(* IEC 61131-3 sources: JingjiangArm/moonboxpro_arm_8.4/Application/Application/任务列表/CommTask/COMM_DIAMONDS/Input_Output, 7 files *)

(* ---- KS_CheckStationOnLine_.st ---- *)
(*@CES
Name=KS_CheckStationOnLine_
Type=FunctionBlock
TypeGuid=6f9dac99-8de1-4efc-8465-68ac443b7d08
Guid=c5e0cdd1-19ab-4cb0-a985-998ee908852c
HasDeclaration=True
HasImplementation=True
*)
{DECLARATION}
FUNCTION KS_CheckStationOnLine_ : BOOL
VAR_INPUT
	i_iSid : INT;
	i_iStationNum : INT;
	i_paiStationId_List : POINTER TO ARRAY [1..128] OF INT;
END_VAR
VAR
	iN : INT;
	xResult : BOOL;
END_VAR

{IMPLEMENTATION}
xResult := FALSE;

FOR iN := 1 TO i_iStationNum BY 1 DO
	IF i_iSid = i_paiStationId_List^[iN] THEN
		xResult := TRUE;
		EXIT;
	END_IF
END_FOR

KS_CheckStationOnLine_ := xResult;

(* ---- KS_Solve_Ver.st ---- *)
(*@CES
Name=KS_Solve_Ver
Type=FunctionBlock
TypeGuid=6f9dac99-8de1-4efc-8465-68ac443b7d08
Guid=eb7c1164-08c4-4977-9280-cbaed44442c1
HasDeclaration=True
HasImplementation=True
*)
{DECLARATION}
FUNCTION KS_Solve_Ver : BOOL(*版本号解析*)
VAR_INPUT
	i_sVersion: STRING;(*版本号*)
	i_pdwYMD: POINTER TO DWORD;
	i_pdwHMS: POINTER TO DWORD;
	i_pdwVer: POINTER TO DWORD;
END_VAR
VAR
END_VAR

{IMPLEMENTATION}
IF i_pdwYMD<>0 AND i_pdwHMS<>0 AND i_pdwVer<>0 THEN

END_IF

(* ---- KS_FB_DIAMONDS_Input.st ---- *)
(*@CES
Name=KS_FB_DIAMONDS_Input
Type=FunctionBlock
TypeGuid=6f9dac99-8de1-4efc-8465-68ac443b7d08
Guid=1e0a50ec-9206-4692-bb5f-e2a5b8087577
HasDeclaration=True
HasImplementation=True
*)
{DECLARATION}
FUNCTION_BLOCK KS_FB_DIAMONDS_Input
VAR_INPUT
	i_xEn: BOOL;
	i_pstStSysParam: POINTER TO StSysParam;
	i_pstStParam_Diamonds_Wr: POINTER TO StParam_Diamonds_Wr;
	i_pstStParam_Diamonds_WrRd: POINTER TO StParam_Diamonds_WrRd;
	i_pstStWrRd_SysCfg: POINTER TO StWrRd_SysCfg;
	i_pstStSysCfgStruct: POINTER TO StSysCfgStruct;
	i_pastStGetMotionSts: POINTER TO ARRAY [1..MAX_STATION_NUM] OF StGetMotionSts;

END_VAR
VAR_OUTPUT
	o_xEn: BOOL;
	o_iErNo: INT;
END_VAR
VAR
	pstStParam_Diamonds_Wr_SysSts : POINTER TO StParam_Diamonds_Wr_SysSts;
	pstStParam_Diamonds_Wr_RdSam : POINTER TO StParam_Diamonds_Wr_RdSam;
	pastStParam_Diamonds_Wr_Err : POINTER TO ARRAY [1..MAX_UNIT_NUM] OF StParam_Diamonds_Wr_Err;
	pastStParam_Diamonds_Wr_RunSts : POINTER TO ARRAY [1..MAX_STATION_NUM] OF StParam_Diamonds_Wr_RunSts;
	iGrp: INT;
	iUnitId: INT;
	byCurSignal_RGB: BYTE;
	abySignalFlag: ARRAY [1..4] OF BYTE;
	iIndex:INT:= 1;
	iN: INT;
	iJ: INT;
	iK: INT;

	abyLastIndex: ARRAY [1..MAX_UNIT_NUM] OF BYTE;
	iAxisId_If: INT;
	iAxisId_Of: INT;
	iGrpId_Uw: INT;
	iGrpId_Rw: INT;
	fbKS_FB_DIAMONDS_SysCfg_WrRd: KS_FB_DIAMONDS_SysCfg_WrRd;
	iMachanicalTypeId: INT;

	astStParam_Diamonds_Wr_RunSts : ARRAY [1..MAX_STATION_NUM] OF StParam_Diamonds_Wr_RunSts;
	iNumIndex: INT:=0;
	iAxisId_T: INT;
	iTypeId_T: INT;
	iUnitId_T: INT;
	iCoreId_T: INT;
	iGroupId_T: INT;
	iAdjAxisId_T: INT;

END_VAR

{IMPLEMENTATION}
o_xEn:= i_xEn;
o_iErNo:= 0;
IF i_xEn THEN
	IF i_pstStSysParam<>0 AND
		i_pstStParam_Diamonds_Wr<>0 AND
		i_pstStParam_Diamonds_WrRd<>0 THEN
		pstStParam_Diamonds_Wr_SysSts:= ADR(i_pstStParam_Diamonds_Wr^.stStParam_Diamonds_Wr_SysSts);
		pstStParam_Diamonds_Wr_RdSam:= ADR(i_pstStParam_Diamonds_Wr^.stStParam_Diamonds_Wr_RdSam);
		pastStParam_Diamonds_Wr_Err:= ADR(i_pstStParam_Diamonds_Wr^.astStParam_Diamonds_Wr_Err);
		pastStParam_Diamonds_Wr_RunSts:= ADR(i_pstStParam_Diamonds_Wr^.astStParam_Diamonds_Wr_RunSts);

		Action_Input_Wr();
(*2025.8.6.195943*)
//2026.5.29.145241		Action_Input_WrRd();

		o_iErNo:= 1;
	ELSE
		o_iErNo:= -2;
	END_IF
ELSE
	o_iErNo:= -1;
END_IF

(* ---- KS_FB_DIAMONDS_Input_WRRD.st ---- *)
(*@CES
Name=KS_FB_DIAMONDS_Input_WRRD
Type=FunctionBlock
TypeGuid=6f9dac99-8de1-4efc-8465-68ac443b7d08
Guid=edee9bc0-245c-42df-bd06-57a10449e106
HasDeclaration=True
HasImplementation=True
*)
{DECLARATION}
FUNCTION_BLOCK KS_FB_DIAMONDS_Input_WRRD
VAR_INPUT
	i_xEn: BOOL;
	i_pstStSysParam: POINTER TO StSysParam;
	i_pstStParam_Diamonds_WrRd: POINTER TO StParam_Diamonds_WrRd;
	i_pstStWrRd_SysCfg: POINTER TO StWrRd_SysCfg;
	i_pstStSysCfgStruct: POINTER TO StSysCfgStruct;

END_VAR
VAR_OUTPUT
	o_xEn: BOOL;
	o_iErNo: INT;
END_VAR
VAR
	iGrp: INT;
	iUnitId: INT;
	byCurSignal_RGB: BYTE;
	abySignalFlag: ARRAY [1..4] OF BYTE;
	iIndex:INT:= 1;
	iN: INT;
	iJ: INT;
	iK: INT;

	abyLastIndex: ARRAY [1..MAX_UNIT_NUM] OF BYTE;
	iAxisId_If: INT;
	iAxisId_Of: INT;
	iGrpId_Uw: INT;
	iGrpId_Rw: INT;
	fbKS_FB_DIAMONDS_SysCfg_WrRd: KS_FB_DIAMONDS_SysCfg_WrRd;
	iMachanicalTypeId: INT;
	iMachanicalTypeId_Tmp: INT;

END_VAR

{IMPLEMENTATION}
(*整机参数|2025.08.06.203301*)
	i_pstStParam_Diamonds_WrRd^.iCustomerId 													:= i_pstStSysParam^.stStSysParam_Save.iCustomerId;									(*客户ID*)
	i_pstStParam_Diamonds_WrRd^.dwEquipmentProf 												:= i_pstStSysParam^.stStSysParam_Save.dwEquipmentProf;								(*设备描述*)
	i_pstStParam_Diamonds_WrRd^.iUnitMaxNum 													:= i_pstStSysParam^.stStSysParam_Save.iUnitMaxNum;												(*最大色组数*)
	i_pstStParam_Diamonds_WrRd^.iCurveViewMaxRange 												:= i_pstStSysParam^.stStSysParam_Save.iCurveViewMaxRange;							(*误差曲线量程上限*)
	i_pstStParam_Diamonds_WrRd^.iTitleTextHeight 												:= i_pstStSysParam^.stStSysParam_Save.iTitleTextHeight;								(*标题字体高度*)
	i_pstStParam_Diamonds_WrRd^.iEntryTextHeight 												:= i_pstStSysParam^.stStSysParam_Save.iEntryTextHeight;								(*输入框字体高度*)
	i_pstStParam_Diamonds_WrRd^.iLabelTextHeight 												:= i_pstStSysParam^.stStSysParam_Save.iLabelTextHeight;								(*标签字体高度*)
	i_pstStParam_Diamonds_WrRd^.iButtonTextHeight 												:= i_pstStSysParam^.stStSysParam_Save.iButtonTextHeight ;							(*按钮字体高度*)
	i_pstStParam_Diamonds_WrRd^.iMessageTextHeight 												:= i_pstStSysParam^.stStSysParam_Save.iMessageTextHeight;							(*消息字体高度*)
	i_pstStParam_Diamonds_WrRd^.byLanguageId 													:= i_pstStSysParam^.stStSysParam_Save.byLanguageId;									(*语言设置*)
	i_pstStParam_Diamonds_WrRd^.byMinutes_ScrSaver 												:= i_pstStSysParam^.stStSysParam_Save.byMinutes_ScrSaver;							(*屏保延时*)
	i_pstStParam_Diamonds_WrRd^.wMachineArchitectureRef 										:= i_pstStSysParam^.stStSysParam_Save.wMachineArchitectureRef;						(*机器架构描述*)
	i_pstStParam_Diamonds_WrRd^.iPromptMsgId 													:= i_pstStSysParam^.stStSysParam_Save.iPromptMsgId;									(*提示信息ID（报警代码）*)
	i_pstStParam_Diamonds_WrRd^.byHorzCtlMode 													:= i_pstStSysParam^.stStSysParam_Save.byHorzCtlMode;								(*横向控制方式-同步-步进-伺服*)
	i_pstStParam_Diamonds_WrRd^.byCheckTimeToTips_BrakeResistance 								:= i_pstStSysParam^.stStSysParam_Save.byCheckTimeToTips_BrakeResistance;			(*制动电阻访问超限提示时间*)
	i_pstStParam_Diamonds_WrRd^.byCheckTimeToEStop_BrakeResistance 								:= i_pstStSysParam^.stStSysParam_Save.byCheckTimeToEStop_BrakeResistance;			(*制动电阻访问超限急停时间*)
	i_pstStParam_Diamonds_WrRd^.byAccessTimes_BrakeResistance 									:= i_pstStSysParam^.stStSysParam_Save.byAccessTimes_BrakeResistance;				(*制动电阻报警限制*)
	i_pstStParam_Diamonds_WrRd^.byAlarmHold_VOL_Uw 												:= i_pstStSysParam^.stStSysParam_Save.byAlarmHold_VOL_Uw;							(*放料没料响应时间*)
	i_pstStParam_Diamonds_WrRd^.byAlarmHold_PrnLength 											:= i_pstStSysParam^.stStSysParam_Save.byAlarmHold_PrnLength;						(*收料印长报警响应时间*)
	i_pstStParam_Diamonds_WrRd^.byHeatingOutWay_III 											:= i_pstStSysParam^.stStSysParam_Save.byHeatingOutWay_III;							(*三档调整方式-只调最低档、只调最高档、三档同时调*)
	i_pstStParam_Diamonds_WrRd^.byHeatingMode 													:= i_pstStSysParam^.stStSysParam_Save.byHeatingMode;								(*温控设置方式切换*)
	i_pstStParam_Diamonds_WrRd^.rOpenThr_Ele 													:= i_pstStSysParam^.stStSysParam_Save.rOpenThr_Ele;									(*电加热开启*)
	i_pstStParam_Diamonds_WrRd^.rCloseThr_Ele 													:= i_pstStSysParam^.stStSysParam_Save.rCloseThr_Ele;								(*电加热关闭*)
	i_pstStParam_Diamonds_WrRd^.rDealValue_Water 												:= i_pstStSysParam^.stStSysParam_Save.rDealValue_Water;								(*水加热死区*)
	i_pstStParam_Diamonds_WrRd^.iMaxOutValue 													:= i_pstStSysParam^.stStSysParam_Save.iMaxOutValue;									(*最大输出*)
	i_pstStParam_Diamonds_WrRd^.iHeatingDebugValue_Water 										:= i_pstStSysParam^.stStSysParam_Save.iHeatingDebugValue_Water;						(*测试开度*)
	i_pstStParam_Diamonds_WrRd^.rKp 															:= i_pstStSysParam^.stStSysParam_Save.rKp;											(*KP*)
	i_pstStParam_Diamonds_WrRd^.rKi 															:= i_pstStSysParam^.stStSysParam_Save.rKi;											(*KI*)
	i_pstStParam_Diamonds_WrRd^.rKd 															:= i_pstStSysParam^.stStSysParam_Save.rKd;											(*Kd*)
	i_pstStParam_Diamonds_WrRd^.iTime_Thres_Water 												:= i_pstStSysParam^.stStSysParam_Save.iTime_Thres_Water;							(*阀门打开时间*)
	i_pstStParam_Diamonds_WrRd^.iCofe_TempCtl_30 												:= i_pstStSysParam^.stStSysParam_Save.iCofe_TempCtl_30;								(*控制阈值1*)
	i_pstStParam_Diamonds_WrRd^.iCofe_TempCtl_30_10 											:= i_pstStSysParam^.stStSysParam_Save.iCofe_TempCtl_30_10;							(*控制阈值2*)
	i_pstStParam_Diamonds_WrRd^.iCofe_TempCtl_10_5 												:= i_pstStSysParam^.stStSysParam_Save.iCofe_TempCtl_10_5;							(*控制阈值3*)
	i_pstStParam_Diamonds_WrRd^.iCofe_TempCtl_5 												:= i_pstStSysParam^.stStSysParam_Save.iCofe_TempCtl_5;								(*控制阈值4*)
	i_pstStParam_Diamonds_WrRd^.iWaterValue_Threshold 											:= i_pstStSysParam^.stStSysParam_Save.iWaterValue_Threshold;						(*水电阈值*)
	i_pstStParam_Diamonds_WrRd^.uiInitDiam_Uw 													:= i_pstStSysParam^.stStSysParam_Save.uiInitDiam_Uw;								(*放料初始卷径*)
	i_pstStParam_Diamonds_WrRd^.uiInitDiam_Rw 													:= i_pstStSysParam^.stStSysParam_Save.uiInitDiam_Rw;								(*收料初始卷径*)
	i_pstStParam_Diamonds_WrRd^.diStepDriveDebugPulse 											:= i_pstStSysParam^.stStSysParam_Save.diStepDriveDebugPulse;						(*测试脉冲数*)
	i_pstStParam_Diamonds_WrRd^.rStepDriveDebugPulse_PosAct 									:= i_pstStSysParam^.stStSysParam_Save.rStepDriveDebugPulse_PosAct;					(*测试距离*)
	i_pstStParam_Diamonds_WrRd^.iStepDriveDebugNum 												:= i_pstStSysParam^.stStSysParam_Save.iStepDriveDebugNum;							(*测试色组号*)
	i_pstStParam_Diamonds_WrRd^.rStepDrivePosPPulse 											:= i_pstStSysParam^.stStSysParam_Save.rStepDrivePosPPulse;							(*单位脉冲距离*)
	i_pstStParam_Diamonds_WrRd^.iStepDrivePulsePRev 											:= i_pstStSysParam^.stStSysParam_Save.iStepDrivePulsePRev;							(*每圈脉冲数*)
	i_pstStParam_Diamonds_WrRd^.iStepDriveSa_Vel 												:= i_pstStSysParam^.stStSysParam_Save.iStepDriveSa_Vel;								(*启动速度*)
	i_pstStParam_Diamonds_WrRd^.iStepDrivePreReg_Vel 											:= i_pstStSysParam^.stStSysParam_Save.iStepDrivePreReg_Vel;							(*预套准速度*)
	i_pstStParam_Diamonds_WrRd^.iStepDriveManu_Vel 												:= i_pstStSysParam^.stStSysParam_Save.iStepDriveManu_Vel;							(*手动低速*)
	i_pstStParam_Diamonds_WrRd^.iStepDriveManu_Vel_Fast 										:= i_pstStSysParam^.stStSysParam_Save.iStepDriveManu_Vel_Fast;						(*手动高速*)
	i_pstStParam_Diamonds_WrRd^.iStepDriveAuto_Vel 												:= i_pstStSysParam^.stStSysParam_Save.iStepDriveAuto_Vel;							(*自动速度*)
	i_pstStParam_Diamonds_WrRd^.iStepDriveAccTime 												:= i_pstStSysParam^.stStSysParam_Save.iStepDriveAccTime;							(*升速时间*)
	i_pstStParam_Diamonds_WrRd^.rHz_MainExhaust_ManuallySet 									:= i_pstStSysParam^.stStSysParam_Save.rHz_MainExhaust_ManuallySet;					(*主排风设定频率*)
	i_pstStParam_Diamonds_WrRd^.byFreq_I_ExhaustAir 											:= i_pstStSysParam^.stStSysParam_Save.byFreq_I_ExhaustAir;							(*排风一档频率*)
	i_pstStParam_Diamonds_WrRd^.byFreq_II_ExhaustAir 											:= i_pstStSysParam^.stStSysParam_Save.byFreq_II_ExhaustAir;							(*排风二档频率*)
	i_pstStParam_Diamonds_WrRd^.byFreq_III_ExhaustAir 											:= i_pstStSysParam^.stStSysParam_Save.byFreq_III_ExhaustAir;						(*排风三档频率*)
	(*待补充-开始|2025.08.06.210116*)
	i_pstStParam_Diamonds_WrRd^.stBitStWrRd_Switch_Machine.xSwitch_PreHotEn_Print				:= i_pstStSysParam^.stStSysParam_Save.xSwitch_PreHotEn_Print				;(*预热印刷激活开关*)
	i_pstStParam_Diamonds_WrRd^.stBitStWrRd_Switch_Machine.xSwitch_ExhAir_Limit_HotWind			:= i_pstStSysParam^.stStSysParam_Save.xSwitch_ExhAir_Limit_HotWind			;(*排风限制热风开关*)
	i_pstStParam_Diamonds_WrRd^.stBitStWrRd_Switch_Machine.xSwitch_ExhAir_Limit_Run				:= i_pstStSysParam^.stStSysParam_Save.xSwitch_ExhAir_Limit_Run				;(*排风限制开机开关*)
	i_pstStParam_Diamonds_WrRd^.stBitStWrRd_Switch_Machine.xSwitch_CommEn_WatchDevice_Tcp		:= i_pstStSysParam^.stStSysParam_Save.xSwitch_CommEn_WatchDevice_Tcp		;(*TCP-外部监控设备开关*)
	i_pstStParam_Diamonds_WrRd^.stBitStWrRd_Switch_Machine.xSwitch_CommEn_WatchDevice_485		:= i_pstStSysParam^.stStSysParam_Save.xSwitch_CommEn_WatchDevice_485		;(*485-外部监控设备开关*)
	i_pstStParam_Diamonds_WrRd^.stBitStWrRd_Switch_Machine.xSwitch_CommEn_1U_485				:= i_pstStSysParam^.stStSysParam_Save.xSwitch_CommEn_1U_485				    ;(*1色人机通讯开关*)
	i_pstStParam_Diamonds_WrRd^.stBitStWrRd_Switch_Machine.xSwitch_CommEn_485					:= i_pstStSysParam^.stStSysParam_Save.xSwitch_CommEn_485					;(*485通讯开关*)
	i_pstStParam_Diamonds_WrRd^.stBitStWrRd_Switch_Machine.xSwitch_CommEn_485_Exh				:= i_pstStSysParam^.stStSysParam_Save.xSwitch_CommEn_485_Exh				;(*排风485通讯开关*)
	i_pstStParam_Diamonds_WrRd^.stBitStWrRd_Switch_Machine.xSwitch_CommEn_485_Scraper			:= i_pstStSysParam^.stStSysParam_Save.xSwitch_CommEn_485_Scraper			;(*刮刀485通讯开关*)
	i_pstStParam_Diamonds_WrRd^.stBitStWrRd_Switch_Machine.xSwitch_CommEn_485_InkRoller			:= i_pstStSysParam^.stStSysParam_Save.xSwitch_CommEn_485_InkRoller			;(*递墨辊485通讯开关*)
	i_pstStParam_Diamonds_WrRd^.stBitStWrRd_Switch_Machine.xSwitch_CommEn_485_HotWind			:= i_pstStSysParam^.stStSysParam_Save.xSwitch_CommEn_485_HotWind			;(*热风485通讯开关*)
	i_pstStParam_Diamonds_WrRd^.stBitStWrRd_Switch_Machine.xSwitch_ArcIntensityBtn_Hmi			:= i_pstStSysParam^.stStSysParam_Save.xSwitch_ArcIntensityBtn_Hmi			;(*手动调节随速度走开关*)
	i_pstStParam_Diamonds_WrRd^.stBitStWrRd_Switch_Machine.xSwitch_PrnRatioIndividual_Setting	:= i_pstStSysParam^.stStSysParam_Save.xSwitch_PrnRatioIndividual_Setting	;(*色组版辊减速比单独设置开关*)
	i_pstStParam_Diamonds_WrRd^.stBitStWrRd_Switch_Machine.xSwitch_NetRatioIndividual_Setting	:= i_pstStSysParam^.stStSysParam_Save.xSwitch_NetRatioIndividual_Setting	;(*色组网辊减速比单独设置开关*)
	i_pstStParam_Diamonds_WrRd^.stBitStWrRd_Switch_Machine.xSwitch_BottomRatioIndividual_Setting:= i_pstStSysParam^.stStSysParam_Save.xSwitch_BottomRatioIndividual_Setting ;(*色组底辊减速比单独设置开关*)
	i_pstStParam_Diamonds_WrRd^.stBitStWrRd_Switch_Machine.xSwitch_StepDriveDebugRun			:= i_pstStSysParam^.stStSysParam_Save.xSwitch_StepDriveDebugRun			    ;(*横向步进电机测试执行开关*)

	i_pstStParam_Diamonds_WrRd^.stBitStWrRd_Switch_Machine.xSetProPointEn					 := i_pstStSysParam^.stStSysParam_Save.xSetProPointEn					;
	i_pstStParam_Diamonds_WrRd^.stBitStWrRd_Switch_Machine.xUseMaxTimeAsSBegin_InLowSpeed    := i_pstStSysParam^.stStSysParam_Save.xUseMaxTimeAsSBegin_InLowSpeed	;
	i_pstStParam_Diamonds_WrRd^.stBitStWrRd_Switch_Machine.xPseudoRandomEn                   := i_pstStSysParam^.stStSysParam_Save.xPseudoRandomEn               	;
	i_pstStParam_Diamonds_WrRd^.stBitStWrRd_Switch_Machine.xPseudoRandomStart                := i_pstStSysParam^.stStSysParam_Save.xPseudoRandomStart            	;
	i_pstStParam_Diamonds_WrRd^.stBitStWrRd_Switch_Machine.xEn_RevLimit                      := i_pstStSysParam^.stStSysParam_Save.xEn_RevLimit                  	;
	i_pstStParam_Diamonds_WrRd^.stBitStWrRd_Switch_Machine.xSaveFineSampleData_ToArc         := i_pstStSysParam^.stStSysParam_Save.xSaveFineSampleData_ToArc     	;
	i_pstStParam_Diamonds_WrRd^.stBitStWrRd_Switch_Machine.xReqSetLedFunc                    := i_pstStSysParam^.stStSysParam_Save.xReqSetLedFunc                	;
	i_pstStParam_Diamonds_WrRd^.stBitStWrRd_Switch_Machine.xSetHmiResolution                 := i_pstStSysParam^.stStSysParam_Save.xSetHmiResolution             	;
	i_pstStParam_Diamonds_WrRd^.stBitStWrRd_Switch_Machine.xPopupWindowVisible               := i_pstStSysParam^.stStSysParam_Save.xPopupWindowVisible           	;
	i_pstStParam_Diamonds_WrRd^.stBitStWrRd_Switch_Machine.xInitArcErr_AjdImmediately        := i_pstStSysParam^.stStSysParam_Save.xInitArcErr_AjdImmediately    	;
	i_pstStParam_Diamonds_WrRd^.stBitStWrRd_Switch_Machine.xPhaseAutoRecoveryEn              := i_pstStSysParam^.stStSysParam_Save.xPhaseAutoRecoveryEn          	;
	i_pstStParam_Diamonds_WrRd^.stBitStWrRd_Switch_Machine.xKeepServo_PreRegisterDne         := i_pstStSysParam^.stStSysParam_Save.xKeepServo_PreRegisterDne     	;
	i_pstStParam_Diamonds_WrRd^.stBitStWrRd_Switch_Machine.xUseIfVel_Uw                      := i_pstStSysParam^.stStSysParam_Save.xUseIfVel_Uw                  	;
	i_pstStParam_Diamonds_WrRd^.stBitStWrRd_Switch_Machine.xKeepServo_Stop                   := i_pstStSysParam^.stStSysParam_Save.xKeepServo_Stop               	;
	i_pstStParam_Diamonds_WrRd^.stBitStWrRd_Switch_Machine.xAxisPrfVelEn                     := i_pstStSysParam^.stStSysParam_Save.xAxisPrfVelEn                 	;
	i_pstStParam_Diamonds_WrRd^.stBitStWrRd_Switch_Machine.xUseGc_PID_2025                   := i_pstStSysParam^.stStSysParam_Save.xUseGc_PID_2025               	;
	i_pstStParam_Diamonds_WrRd^.stBitStWrRd_Switch_Machine.xFlag_Follow_1U_Double_V          := i_pstStSysParam^.stStSysParam_Save.xFlag_Follow_1U_Double_V      	;
	i_pstStParam_Diamonds_WrRd^.stBitStWrRd_Switch_Machine.xArcErrCorrectIsRev_V             := i_pstStSysParam^.stStSysParam_Save.xArcErrCorrectIsRev_V         	;
	i_pstStParam_Diamonds_WrRd^.stBitStWrRd_Switch_Machine.xAutoSetSampleType                := i_pstStSysParam^.stStSysParam_Save.xAutoSetSampleType            	;
	i_pstStParam_Diamonds_WrRd^.stBitStWrRd_Switch_Machine.xGetSampleTypeBtn                 := i_pstStSysParam^.stStSysParam_Save.xGetSampleTypeBtn             	;
	i_pstStParam_Diamonds_WrRd^.stBitStWrRd_Switch_Machine.xAutoSetArcCtlWay                 := i_pstStSysParam^.stStSysParam_Save.xAutoSetArcCtlWay	;
	i_pstStParam_Diamonds_WrRd^.stBitStWrRd_Switch_Machine.xWorkMode_Inch:= i_pstStSysParam^.stStSysParam_Save.xWorkMode_Inch;
	i_pstStParam_Diamonds_WrRd^.stBitStWrRd_Switch_Machine.xSwitch_ScraperReset:= i_pstStSysParam^.stStSysParam_UnSave.xSwitch_ScraperReset;
	i_pstStParam_Diamonds_WrRd^.stBitStWrRd_Switch_Machine.xSwitch_InkRollerReset:= i_pstStSysParam^.stStSysParam_UnSave.xSwitch_InkRollerReset;
	i_pstStParam_Diamonds_WrRd^.stBitStWrRd_Switch_Machine.xSwitch_HotwindReset:= i_pstStSysParam^.stStSysParam_UnSave.xSwitch_HotwindReset;
	i_pstStParam_Diamonds_WrRd^.stBitStWrRd_Switch_Machine.xSwitch_ResetTemctlModule:= i_pstStSysParam^.stStSysParam_UnSave.xSwitch_ResetTemctlModule;
	i_pstStParam_Diamonds_WrRd^.stBitStWrRd_Switch_Machine.xSwitch_Copy1stUExhaustDamperPos:= i_pstStSysParam^.stStSysParam_UnSave.xSwitch_Copy1stUExhaustDamperPos;
	i_pstStParam_Diamonds_WrRd^.stBitStWrRd_Switch_Machine.xMoveFreq_I_ToAll_AirHot:= i_pstStSysParam^.stStSysParam_UnSave.xMoveFreq_I_ToAll_AirHot;
	i_pstStParam_Diamonds_WrRd^.stBitStWrRd_Switch_Machine.xMoveFreq_II_ToAll_AirHot:= i_pstStSysParam^.stStSysParam_UnSave.xMoveFreq_II_ToAll_AirHot;
	i_pstStParam_Diamonds_WrRd^.stBitStWrRd_Switch_Machine.xMoveFreq_III_ToAll_AirHot:= i_pstStSysParam^.stStSysParam_UnSave.xMoveFreq_III_ToAll_AirHot;
	i_pstStParam_Diamonds_WrRd^.stBitStWrRd_Switch_Machine.xMoveFreq_I_ToAll_ExhaustAir:= i_pstStSysParam^.stStSysParam_UnSave.xMoveFreq_I_ToAll_ExhaustAir;
	i_pstStParam_Diamonds_WrRd^.stBitStWrRd_Switch_Machine.xMoveFreq_II_ToAll_ExhaustAir:= i_pstStSysParam^.stStSysParam_UnSave.xMoveFreq_II_ToAll_ExhaustAir;
	i_pstStParam_Diamonds_WrRd^.stBitStWrRd_Switch_Machine.xMoveFreq_III_ToAll_ExhaustAir:= i_pstStSysParam^.stStSysParam_UnSave.xMoveFreq_III_ToAll_ExhaustAir;

	////////////////////////////////////////////////////////////分割线///////////////////////////////////////////////
(*2025.8.25.152610||增加当前波形通道选择2025.8.25.152623*)
	i_pstStParam_Diamonds_WrRd^.iUid_Choose:= i_pstStSysParam^.stStSysParam_Save.iUid		;
	(*待补充-结束|2025.08.06.210116*)
(*2025.10.24.132427*)(*油墨槽控制相关*)
	i_pstStParam_Diamonds_WrRd^.xInkGrooveCtlEn					:= i_pstStSysParam^.stStSysParam_Save.xInkGrooveCtlEn;
	i_pstStParam_Diamonds_WrRd^.xInkGrooveCtlDirRev					:= i_pstStSysParam^.stStSysParam_Save.xInkGrooveCtlDirRev;
	i_pstStParam_Diamonds_WrRd^.xInkGrooveCali_Hmi					:= i_pstStSysParam^.stStSysParam_UnSave.xInkGrooveCali_Hmi;
	i_pstStParam_Diamonds_WrRd^.iInkGroove_Vel					:= i_pstStSysParam^.stStSysParam_Save.iInkGroove_Vel;
	i_pstStParam_Diamonds_WrRd^.iInkGrooveMoveDis_Max					:= i_pstStSysParam^.stStSysParam_Save.iInkGrooveMoveDis_Max;
	i_pstStParam_Diamonds_WrRd^.iInkGrooveSa_Vel					:= i_pstStSysParam^.stStSysParam_Save.iInkGrooveSa_Vel;
	i_pstStParam_Diamonds_WrRd^.iInkGrooveAccTime					:= i_pstStSysParam^.stStSysParam_Save.iInkGrooveAccTime;
	i_pstStParam_Diamonds_WrRd^.iInkGroovePulsePRev					:= i_pstStSysParam^.stStSysParam_Save.iInkGroovePulsePRev;
	i_pstStParam_Diamonds_WrRd^.rInkGroovePosPPulse					:= i_pstStSysParam^.stStSysParam_Save.rInkGroovePosPPulse;
	i_pstStParam_Diamonds_WrRd^.iTimeOut_Slave_485_Inverter			:= i_pstStSysParam^.stStSysParam_Save.iTimeOut_Slave_485_Inverter;
	i_pstStParam_Diamonds_WrRd^.byModbusNum_Max						:= i_pstStSysParam^.stStSysParam_Save.byModbusNum_Max;
	i_pstStParam_Diamonds_WrRd^.byFreq_I_AirHot:= i_pstStSysParam^.stStSysParam_Save.byFreq_I_AirHot;
	i_pstStParam_Diamonds_WrRd^.byFreq_II_AirHot:= i_pstStSysParam^.stStSysParam_Save.byFreq_II_AirHot;
	i_pstStParam_Diamonds_WrRd^.byFreq_III_AirHot:= i_pstStSysParam^.stStSysParam_Save.byFreq_III_AirHot;
	i_pstStParam_Diamonds_WrRd^.byFreq_I_ExhaustAir:= i_pstStSysParam^.stStSysParam_Save.byFreq_I_ExhaustAir;
	i_pstStParam_Diamonds_WrRd^.byFreq_II_ExhaustAir:= i_pstStSysParam^.stStSysParam_Save.byFreq_II_ExhaustAir;
	i_pstStParam_Diamonds_WrRd^.byFreq_III_ExhaustAir:= i_pstStSysParam^.stStSysParam_Save.byFreq_III_ExhaustAir;
(*2025.10.28.112509*)
i_pstStParam_Diamonds_WrRd^.byExhaustMode:= i_pstStSysParam^.stStSysParam_Save.byExhaustMode;
i_pstStParam_Diamonds_WrRd^.byExhaustLinkageNum:= i_pstStSysParam^.stStSysParam_Save.byExhaustLinkageNum;
i_pstStParam_Diamonds_WrRd^.byFreqMax_ExhaustAir:= i_pstStSysParam^.stStSysParam_Save.byFreqMax_ExhaustAir;
i_pstStParam_Diamonds_WrRd^.byFreqMin_ExhaustAir:= i_pstStSysParam^.stStSysParam_Save.byFreqMin_ExhaustAir;
i_pstStParam_Diamonds_WrRd^.byCoefExhaust:= i_pstStSysParam^.stStSysParam_Save.byCoefExhaust;
(*2025.10.28.112715处理一下机械参数*)
//2026.05.26.214359 查漏补缺
i_pstStParam_Diamonds_WrRd^.byOverPercent_RatedRpm:= i_pstStSysParam^.stStSysParam_Save.byOverPercent_RatedRpm;
i_pstStParam_Diamonds_WrRd^.uiMaxDia:= i_pstStSysParam^.stStSysParam_Save.uiMaxDia;

	i_pstStParam_Diamonds_WrRd^.byMachanicalTypeId:= g_stStSysParam.stStSysParam_Save.byMechanicalTypeId;
	iMachanicalTypeId:= BYTE_TO_INT(i_pstStParam_Diamonds_WrRd^.byMachanicalTypeId);
//	IF iMachanicalTypeId>=1 AND iMachanicalTypeId<=5 THEN
	FOR iMachanicalTypeId_Tmp:=1 TO 5 BY 1 DO
		SysMemCpy(
			ADR(i_pstStParam_Diamonds_WrRd^.astStMechanicalParamBuf[iMachanicalTypeId_Tmp].abyBuf),
			ADR(i_pstStSysParam^.stStSysParam_Save.astStMechanicalParamBuf[iMachanicalTypeId_Tmp].abyBuf),
			SIZEOF(i_pstStParam_Diamonds_WrRd^.astStMechanicalParamBuf[iMachanicalTypeId_Tmp].abyBuf),
		);
	END_FOR
//	END_IF
	(*2025.7.3.175755——||| 9905界面参数*)
	i_pstStParam_Diamonds_WrRd^.uiMaxVel_UseCalcAcc							:= i_pstStSysParam^.stStSysParam_Save.uiMaxVel_UseCalcAcc				;
	i_pstStParam_Diamonds_WrRd^.byPseudoRandomRoundTimes					:= i_pstStSysParam^.stStSysParam_Save.byPseudoRandomRoundTimes			;
	i_pstStParam_Diamonds_WrRd^.rPseudoRandomAmplitude						:= i_pstStSysParam^.stStSysParam_Save.rPseudoRandomAmplitude			;
	i_pstStParam_Diamonds_WrRd^.bySetTestPid_IfOf							:= i_pstStSysParam^.stStSysParam_Save.bySetTestPid_IfOf					;
	i_pstStParam_Diamonds_WrRd^.by10vSignalCoef								:= i_pstStSysParam^.stStSysParam_Save.by10vSignalCoef					;
	i_pstStParam_Diamonds_WrRd^.rCompensateGirthWhenAccing_If				:= i_pstStSysParam^.stStSysParam_Save.rCompensateGirthWhenAccing_If		;
	i_pstStParam_Diamonds_WrRd^.rCompensateGirthWhenAccing_Of				:= i_pstStSysParam^.stStSysParam_Save.rCompensateGirthWhenAccing_Of		;
	i_pstStParam_Diamonds_WrRd^.byArcDeCoupleStepTest						:= i_pstStSysParam^.stStSysParam_Save.byArcDeCoupleStepTest				;
	i_pstStParam_Diamonds_WrRd^.iCustomerLogoOffsetX						:= i_pstStSysParam^.stStSysParam_Save.iCustomerLogoOffsetX				;
	i_pstStParam_Diamonds_WrRd^.byGuardrialColor_R							:= i_pstStSysParam^.stStSysParam_Save.byGuardrialColor_R				;
	i_pstStParam_Diamonds_WrRd^.byGuardrialColor_G							:= i_pstStSysParam^.stStSysParam_Save.byGuardrialColor_G				;
	i_pstStParam_Diamonds_WrRd^.byGuardrialColor_B							:= i_pstStSysParam^.stStSysParam_Save.byGuardrialColor_B				;
	i_pstStParam_Diamonds_WrRd^.iLedFuncId									:= i_pstStSysParam^.stStSysParam_Save.iLedFuncId						;
	i_pstStParam_Diamonds_WrRd^.iSetHmiResValue								:= i_pstStSysParam^.stStSysParam_Save.iSetHmiResValue					;
	i_pstStParam_Diamonds_WrRd^.wRunningTime_Day							:= i_pstStSysParam^.stStSysParam_Save.wRunningTime_Day					;
	i_pstStParam_Diamonds_WrRd^.byRunningTime_Hour							:= i_pstStSysParam^.stStSysParam_Save.byRunningTime_Hour				;
	i_pstStParam_Diamonds_WrRd^.byRunningTime_Min							:= i_pstStSysParam^.stStSysParam_Save.byRunningTime_Min					;
	i_pstStParam_Diamonds_WrRd^.byRunningTime_Sec							:= i_pstStSysParam^.stStSysParam_Save.byRunningTime_Sec					;
	i_pstStParam_Diamonds_WrRd^.byArcIntensity_W							:= i_pstStSysParam^.stStSysParam_Save.byArcIntensity_W					;
	i_pstStParam_Diamonds_WrRd^.byArcIntensity_M							:= i_pstStSysParam^.stStSysParam_Save.byArcIntensity_M					;
	i_pstStParam_Diamonds_WrRd^.byArcIntensity_S							:= i_pstStSysParam^.stStSysParam_Save.byArcIntensity_S					;
	i_pstStParam_Diamonds_WrRd^.byMotorOverTempValue_UseEncTemp				:= i_pstStSysParam^.stStSysParam_Save.byMotorOverTempValue_UseEncTemp	;
	i_pstStParam_Diamonds_WrRd^.byRemainSpaceNum_PTCTL         				:= i_pstStSysParam^.stStSysParam_Save.byRemainSpaceNum_PTCTL         	;
	i_pstStParam_Diamonds_WrRd^.rSpeed_SCoeff_Type789          				:= i_pstStSysParam^.stStSysParam_Save.rSpeed_SCoeff_Type789          	;
	i_pstStParam_Diamonds_WrRd^.byMaxPulseOut_16dIO            				:= i_pstStSysParam^.stStSysParam_Save.byMaxPulseOut_16dIO            	;
	i_pstStParam_Diamonds_WrRd^.bySysSamplePrecision           				:= i_pstStSysParam^.stStSysParam_Save.bySysSamplePrecision           	;
	i_pstStParam_Diamonds_WrRd^.byArcAdjValueDealType          				:= i_pstStSysParam^.stStSysParam_Save.byArcAdjValueDealType          	;
	i_pstStParam_Diamonds_WrRd^.byArcErrLimitToCtl_P           				:= i_pstStSysParam^.stStSysParam_Save.byArcErrLimitToCtl_P           	;
	i_pstStParam_Diamonds_WrRd^.byArcErrLimitToCtl_I           				:= i_pstStSysParam^.stStSysParam_Save.byArcErrLimitToCtl_I           	;
	i_pstStParam_Diamonds_WrRd^.byMaxPulseOut_Module           				:= i_pstStSysParam^.stStSysParam_Save.byMaxPulseOut_Module           	;
	i_pstStParam_Diamonds_WrRd^.byArcFineSampleType            				:= i_pstStSysParam^.stStSysParam_Save.byArcFineSampleType            	;
	i_pstStParam_Diamonds_WrRd^.byArcPidGetType                				:= i_pstStSysParam^.stStSysParam_Save.byArcPidGetType                	;
	i_pstStParam_Diamonds_WrRd^.rFilmLenth_Eyes                				:= i_pstStSysParam^.stStSysParam_Save.rFilmLenth_Eyes                	;
	i_pstStParam_Diamonds_WrRd^.uiArcSysDelayTime_ms           				:= i_pstStSysParam^.stStSysParam_Save.uiArcSysDelayTime_ms           	;
	i_pstStParam_Diamonds_WrRd^.byParamIndex_Huang							:= i_pstStSysParam^.stStSysParam_Save.byParamIndex_Huang				;
	i_pstStParam_Diamonds_WrRd^.uiControllerVel_Huang						:= i_pstStSysParam^.stStSysParam_Save.uiControllerVel_Huang				;
	i_pstStParam_Diamonds_WrRd^.byCouplingType								:= i_pstStSysParam^.stStSysParam_Save.byCouplingType					;
	i_pstStParam_Diamonds_WrRd^.byDeCoupleArcNum							:= i_pstStSysParam^.stStSysParam_Save.byDeCoupleArcNum					;

//2026.4.25.144922
	i_pstStParam_Diamonds_WrRd^.byArcIntensity								:= i_pstStSysParam^.stStSysParam_Save.byArcIntensity;

(*系参数|2025.08.06.202852*)
FOR iGrp:=1 TO 2 BY 1 DO
	i_pstStParam_Diamonds_WrRd^.arGirth_AxiaA_Uw[iGrp]  := i_pstStSysParam^.astStGrpParam_Save[iGrp].rGirth_AxiaA_Uw;								(*放料A轴周长*)
	i_pstStParam_Diamonds_WrRd^.arGirth_AxiaB_Uw[iGrp]  := i_pstStSysParam^.astStGrpParam_Save[iGrp].rGirth_AxiaB_Uw ;								(*放料B轴周长*)
	i_pstStParam_Diamonds_WrRd^.arGirth_AxiaA_Rw[iGrp]  := i_pstStSysParam^.astStGrpParam_Save[iGrp].rGirth_AxiaA_Rw ;								(*收料A轴周长*)
	i_pstStParam_Diamonds_WrRd^.arGirth_AxiaB_Rw[iGrp]  := i_pstStSysParam^.astStGrpParam_Save[iGrp].rGirth_AxiaB_Rw ;								(*收料B轴周长*)
	i_pstStParam_Diamonds_WrRd^.arGirth_Pu[iGrp]        := i_pstStSysParam^.astStGrpParam_Save[iGrp].rGirth_PrnRoller ;								(*版周长*)
	i_pstStParam_Diamonds_WrRd^.arTaper_Begin_Rw[iGrp]  := i_pstStSysParam^.astStGrpParam_UnSave[iGrp].rTaperValueBegin_Hmi_Rw ;								(*收料锥度-大张力*)
	i_pstStParam_Diamonds_WrRd^.arTaper_End_Rw[iGrp]    := i_pstStSysParam^.astStGrpParam_UnSave[iGrp].rTaperValueEnd_Hmi_Rw ;								(*收料锥度-小张力*)
	i_pstStParam_Diamonds_WrRd^.arVel_Tar[iGrp]         := i_pstStSysParam^.astStGrpParam_Save[iGrp].rVel_Tar ;										(*目标速度*)
	i_pstStParam_Diamonds_WrRd^.aiTime_AutoAcc[iGrp]    := i_pstStSysParam^.astStGrpParam_Save[iGrp].iTime_AutoAcc ;								(*自动加速时间（S）*)
	i_pstStParam_Diamonds_WrRd^.aiTime_AutoDec[iGrp]    := i_pstStSysParam^.astStGrpParam_Save[iGrp].iTime_AutoDec ;								(*自动减速时间（S）*)
	i_pstStParam_Diamonds_WrRd^.aiTime_ManuAcc[iGrp]    := i_pstStSysParam^.astStGrpParam_Save[iGrp].iTime_ManuAcc ;								(*手动加速时间（S）*)
	i_pstStParam_Diamonds_WrRd^.aiTime_ManuDec[iGrp]    := i_pstStSysParam^.astStGrpParam_Save[iGrp].iTime_ManuDec ;								(*手动减速时间（S）*)
	i_pstStParam_Diamonds_WrRd^.aiTime_FastStop[iGrp]   := i_pstStSysParam^.astStGrpParam_Save[iGrp].iTime_FastStop ;								(*快停时间（S）*)
	i_pstStParam_Diamonds_WrRd^.aiTime_Estop[iGrp]      := i_pstStSysParam^.astStGrpParam_Save[iGrp].iTime_Estop ;									(*急停时间（S)*)
	i_pstStParam_Diamonds_WrRd^.aiTime_Stop[iGrp]      := i_pstStSysParam^.astStGrpParam_Save[iGrp].iTime_Stop ;									(*急停时间（S)*)
	i_pstStParam_Diamonds_WrRd^.adwPrnLen_Alarm[iGrp,1]:= LREAL_TO_DWORD(i_pstStSysParam^.astStGrpParam_Save[iGrp].alrPrnLen_Alr[1]);								(*印长报警*)
	i_pstStParam_Diamonds_WrRd^.adwPrnLen_Alarm[iGrp,2]:= LREAL_TO_DWORD(i_pstStSysParam^.astStGrpParam_Save[iGrp].alrPrnLen_Alr[2]);								(*印长报警*)
	i_pstStParam_Diamonds_WrRd^.adwPrnLen_Alarm[iGrp,3]:= LREAL_TO_DWORD(i_pstStSysParam^.astStGrpParam_Save[iGrp].alrPrnLen_Alr[3]);								(*印长报警*)
	(*待补充-开始|2025.08.06.215021*)
	i_pstStParam_Diamonds_WrRd^.astBitStWrRd_Switch_Grp[iGrp].xSwitch_MachineRev			:= i_pstStSysParam^.astStGrpParam_UnSave[iGrp].xMachineRev 	;(*反向走料开关*)
	i_pstStParam_Diamonds_WrRd^.astBitStWrRd_Switch_Grp[iGrp].xSwitch_6Inch_Rw				:= i_pstStSysParam^.astStGrpParam_Save[iGrp].xUseKnob_6Inch_Rw_Hmi 	;(*收料3/6吋选择开关*)
	i_pstStParam_Diamonds_WrRd^.astBitStWrRd_Switch_Grp[iGrp].xSwitch_StartUp				:= i_pstStSysParam^.astStGrpParam_Save[iGrp].xSwitch_StartUp 	;(*一键开机开关*)
	i_pstStParam_Diamonds_WrRd^.astBitStWrRd_Switch_Grp[iGrp].xSwitch_DiamMeasureAuto		:= i_pstStSysParam^.astStGrpParam_Save[iGrp].xDiamMeasureAutomatic_Uw 	;(*自动卷径开关*)
	i_pstStParam_Diamonds_WrRd^.astBitStWrRd_Switch_Grp[iGrp].xSwitch_RollOver				:= i_pstStSysParam^.astStGrpParam_Save[iGrp].xSwitch_RollOver	;(*设备翻料架开关*)
	i_pstStParam_Diamonds_WrRd^.astBitStWrRd_Switch_Grp[iGrp].xSwitch_Thickness				:= i_pstStSysParam^.astStGrpParam_Save[iGrp].xGetFilmThickNessAuto 	;(*料膜厚度手自动获取开关*)
	i_pstStParam_Diamonds_WrRd^.astBitStWrRd_Switch_Grp[iGrp].xSwitch_CutDneResetPidEn_Uw	:= i_pstStSysParam^.astStGrpParam_Save[iGrp].xCutDneResetPidEn_Uw 	;(*放料裁切后系数手自动*)
	i_pstStParam_Diamonds_WrRd^.astBitStWrRd_Switch_Grp[iGrp].xSwitch_CutDneResetPidEn_Rw	:= i_pstStSysParam^.astStGrpParam_Save[iGrp].xCutDneResetPidEn_Rw 	;(*收料裁切后系数手自动*)
	i_pstStParam_Diamonds_WrRd^.astBitStWrRd_Switch_Grp[iGrp].xSwitch_AutomaticCutEn_Uw		:= i_pstStSysParam^.astStGrpParam_Save[iGrp].xAutomaticCutEn_Uw 	;(*放料自动接料是能*)
	i_pstStParam_Diamonds_WrRd^.astBitStWrRd_Switch_Grp[iGrp].xSwitch_AutomaticCutEn_Rw		:= i_pstStSysParam^.astStGrpParam_Save[iGrp].xAutomaticCutEn_Rw 	;(*放料自动接料是能*)
	i_pstStParam_Diamonds_WrRd^.astBitStWrRd_Switch_Grp[iGrp].xSwitch_AutoAdjust_V_Grp		:= i_pstStSysParam^.astStGrpParam_UnSave[iGrp].xSwitch_AutoAdjust_V_Grp 	;(*整机纵向自动调整开关*)
	i_pstStParam_Diamonds_WrRd^.astBitStWrRd_Switch_Grp[iGrp].xSwitch_AutoAdjust_H_Grp		:= i_pstStSysParam^.astStGrpParam_UnSave[iGrp].xSwitch_AutoAdjust_H_Grp 	;(*整机纵向自动调整开关*)
	i_pstStParam_Diamonds_WrRd^.astBitStWrRd_Switch_Grp[iGrp].xSwitch_Follow_1U_V_Grp		:= i_pstStSysParam^.astStGrpParam_Save[iGrp].xFlag_Follow_1U_V 	;(*纵向跟1色开关*)
	i_pstStParam_Diamonds_WrRd^.astBitStWrRd_Switch_Grp[iGrp].xSwitch_Follow_1U_H_Grp		:= i_pstStSysParam^.astStGrpParam_Save[iGrp].xFlag_Follow_1U_H 	;(*横向跟1色开关*)
	i_pstStParam_Diamonds_WrRd^.astBitStWrRd_Switch_Grp[iGrp].xSwitch_DiamAuto_Pot			:= i_pstStSysParam^.astStGrpParam_Save[iGrp].byDiamMeasureTypeId_Uw=1 	;(*卷径检测使用电位器*)
	i_pstStParam_Diamonds_WrRd^.astBitStWrRd_Switch_Grp[iGrp].xSwitch_DiamAuto_Enc			:= i_pstStSysParam^.astStGrpParam_Save[iGrp].byDiamMeasureTypeId_Uw=2 	;(*卷径检测使用编码器*)
	i_pstStParam_Diamonds_WrRd^.astBitStWrRd_Switch_Grp[iGrp].xSwitch_DiamAuto_Ultrasonic_S	:= i_pstStSysParam^.astStGrpParam_Save[iGrp].byDiamMeasureTypeId_Uw=3 	;(*卷径检测使用单超声波*)
	i_pstStParam_Diamonds_WrRd^.astBitStWrRd_Switch_Grp[iGrp].xSwitch_DiamAuto_Ultrasonic_D	:= i_pstStSysParam^.astStGrpParam_Save[iGrp].byDiamMeasureTypeId_Uw=4 	;(*卷径检测使用双超声波*)
	i_pstStParam_Diamonds_WrRd^.astBitStWrRd_Switch_Grp[iGrp].xSwitch_DiamAuto_DualParam	:= i_pstStSysParam^.astStGrpParam_Save[iGrp].xFlag_AxisABParaFroDiaMea_Uw 	;(*卷径检测双轴参数分开*)
	i_pstStParam_Diamonds_WrRd^.astBitStWrRd_Switch_Grp[iGrp].xSwitch_DebugMode				:= i_pstStSysParam^.astStGrpParam_UnSave[iGrp].xIsDebugMode_Machine 	;(*调试模式开关*)
	i_pstStParam_Diamonds_WrRd^.astBitStWrRd_Switch_Grp[iGrp].xSwitch_Debug_DiamMeasure_Uw	:= i_pstStSysParam^.astStGrpParam_UnSave[iGrp].xIsDebug_DiaMeasure_Uw 	;(*放料卷径检测电位器调试开关*)
	i_pstStParam_Diamonds_WrRd^.astBitStWrRd_Switch_Grp[iGrp].xBtn_Diameasure_Confirm_1		:= i_pstStSysParam^.astStGrpParam_UnSave[iGrp].axMeasure_StdVol[1] 	;(*自动卷径标定——1*)
	i_pstStParam_Diamonds_WrRd^.astBitStWrRd_Switch_Grp[iGrp].xBtn_Diameasure_Confirm_2		:= i_pstStSysParam^.astStGrpParam_UnSave[iGrp].axMeasure_StdVol[2] 	;(*自动卷径标定——2*)
	i_pstStParam_Diamonds_WrRd^.astBitStWrRd_Switch_Grp[iGrp].xBtn_Diameasure_Confirm_3		:= i_pstStSysParam^.astStGrpParam_UnSave[iGrp].axMeasure_StdVol[3]	;(*自动卷径标定——3*)
	i_pstStParam_Diamonds_WrRd^.astBitStWrRd_Switch_Grp[iGrp].xBtn_Diameasure_Confirm_4		:= i_pstStSysParam^.astStGrpParam_UnSave[iGrp].axMeasure_StdVol[4]	;(*自动卷径标定——4*)
	i_pstStParam_Diamonds_WrRd^.astBitStWrRd_Switch_Grp[iGrp].xSwitch_CutUseReflectionSensor				:= i_pstStSysParam^.astStGrpParam_Save[iGrp].xCutUseReflectionSensor_Uw ;(*放料裁切使用弧面开关*)
	i_pstStParam_Diamonds_WrRd^.astBitStWrRd_Switch_Grp[iGrp].xSwitch_UseAbsEnc_Uw				:= i_pstStSysParam^.astStGrpParam_Save[iGrp].xUseAbsEncoder_Uw					;(*放料使用绝对值编码器开关*)
	i_pstStParam_Diamonds_WrRd^.astBitStWrRd_Switch_Grp[iGrp].xSwitch_AxisLocaltion_DualParam_Uw	:= i_pstStSysParam^.astStGrpParam_Save[iGrp].xEn_DualParam_AbsEncLocation_Uw	;(*放料绝对值编码器定位双轴参数开关*)
	i_pstStParam_Diamonds_WrRd^.astBitStWrRd_Switch_Grp[iGrp].xSwitch_Debug_Axis_Uw				:= i_pstStSysParam^.astStGrpParam_UnSave[iGrp].xDebug_Enc_Uw					;(*放料轴运行调试模式*)
	i_pstStParam_Diamonds_WrRd^.astBitStWrRd_Switch_Grp[iGrp].xSwitch_Debug_Uw_CutUpChoose		:= i_pstStSysParam^.astStGrpParam_UnSave[iGrp].xCutterOnTopFroDebug_Uw			;(*放料绝对值编码器定位调试-上裁选择*)
	i_pstStParam_Diamonds_WrRd^.astBitStWrRd_Switch_Grp[iGrp].xSwitch_Debug_Uw_AxisA_Choose		:= i_pstStSysParam^.astStGrpParam_UnSave[iGrp].xCurAxisAFroDebug_Uw			;

	i_pstStParam_Diamonds_WrRd^.astBitStWrRd_Switch_Grp[iGrp].xSwitch_UseAbsEnc_Rw				:= i_pstStSysParam^.astStGrpParam_Save[iGrp].xUseAbsEncoder_Rw					;(*放料使用绝对值编码器开关*)
	i_pstStParam_Diamonds_WrRd^.astBitStWrRd_Switch_Grp[iGrp].xSwitch_AxisLocaltion_DualParam_Rw	:= i_pstStSysParam^.astStGrpParam_Save[iGrp].xSwitch_AxisLocaltion_DualParam_Rw;
	i_pstStParam_Diamonds_WrRd^.astBitStWrRd_Switch_Grp[iGrp].xSwitch_Debug_Axis_Rw				:= i_pstStSysParam^.astStGrpParam_UnSave[iGrp].xDebug_Enc_Rw					;
	i_pstStParam_Diamonds_WrRd^.astBitStWrRd_Switch_Grp[iGrp].xSwitch_Debug_Rw_CutUpChoose		:= i_pstStSysParam^.astStGrpParam_UnSave[iGrp].xCutterOnTopFroDebug_Rw			;(*放料绝对值编码器定位调试-上裁选择*)
	i_pstStParam_Diamonds_WrRd^.astBitStWrRd_Switch_Grp[iGrp].xSwitch_Debug_Rw_AxisA_Choose		:= i_pstStSysParam^.astStGrpParam_UnSave[iGrp].xCurAxisAFroDebug_Rw			;
	i_pstStParam_Diamonds_WrRd^.astBitStWrRd_Switch_Grp[iGrp].xSwitch_Scrap_Avoidance:= i_pstStSysParam^.astStGrpParam_Save[iGrp].xSwitch_GiveupHeaderEn;
	i_pstStParam_Diamonds_WrRd^.astBitStWrRd_Switch_Grp[iGrp].xSwitch_CCW_AfterCut_Uw:= i_pstStSysParam^.astStGrpParam_Save[iGrp].xFlag_CCW_AfterCutted_Uw;
	i_pstStParam_Diamonds_WrRd^.astBitStWrRd_Switch_Grp[iGrp].xSwitch_UseRadCompensate_Uw:= i_pstStSysParam^.astStGrpParam_Save[iGrp].xUseRadCompensate_Uw;
	i_pstStParam_Diamonds_WrRd^.astBitStWrRd_Switch_Grp[iGrp].xSwitch_TowerDir_Uw:= i_pstStSysParam^.astStGrpParam_Save[iGrp].xTowerDir_Uw;
	i_pstStParam_Diamonds_WrRd^.astBitStWrRd_Switch_Grp[iGrp].xSwitch_Debug_Spd_Uw:= i_pstStSysParam^.astStGrpParam_UnSave[iGrp].wAxisDebug_UwRw.0;
	i_pstStParam_Diamonds_WrRd^.astBitStWrRd_Switch_Grp[iGrp].xBtn_DebugSpdAxisA_Uw_MoveEn	:=i_pstStSysParam^.astStGrpParam_UnSave[iGrp].wAxisDebug_UwRw.1;
	i_pstStParam_Diamonds_WrRd^.astBitStWrRd_Switch_Grp[iGrp].xBtn_DebugSpdAxisA_Uw_AccEn	:=i_pstStSysParam^.astStGrpParam_UnSave[iGrp].wAxisDebug_UwRw.2;
	i_pstStParam_Diamonds_WrRd^.astBitStWrRd_Switch_Grp[iGrp].xBtn_DebugSpdAxisB_Uw_MoveEn	:=i_pstStSysParam^.astStGrpParam_UnSave[iGrp].wAxisDebug_UwRw.4;
	i_pstStParam_Diamonds_WrRd^.astBitStWrRd_Switch_Grp[iGrp].xBtn_DebugSpdAxisB_Uw_AccEn	:=i_pstStSysParam^.astStGrpParam_UnSave[iGrp].wAxisDebug_UwRw.5;
	i_pstStParam_Diamonds_WrRd^.astBitStWrRd_Switch_Grp[iGrp].xSwitch_Debug_Spd_Rw:= i_pstStSysParam^.astStGrpParam_UnSave[iGrp].wAxisDebug_UwRw.8;
	i_pstStParam_Diamonds_WrRd^.astBitStWrRd_Switch_Grp[iGrp].xBtn_DebugSpdAxisA_Rw_MoveEn	:= i_pstStSysParam^.astStGrpParam_UnSave[iGrp].wAxisDebug_UwRw.9;
	i_pstStParam_Diamonds_WrRd^.astBitStWrRd_Switch_Grp[iGrp].xBtn_DebugSpdAxisA_Rw_AccEn	:= i_pstStSysParam^.astStGrpParam_UnSave[iGrp].wAxisDebug_UwRw.10;
	i_pstStParam_Diamonds_WrRd^.astBitStWrRd_Switch_Grp[iGrp].xBtn_DebugSpdAxisB_Rw_MoveEn	:= i_pstStSysParam^.astStGrpParam_UnSave[iGrp].wAxisDebug_UwRw.12;
	i_pstStParam_Diamonds_WrRd^.astBitStWrRd_Switch_Grp[iGrp].xBtn_DebugSpdAxisB_Rw_AccEn	:= i_pstStSysParam^.astStGrpParam_UnSave[iGrp].wAxisDebug_UwRw.13;
 	i_pstStParam_Diamonds_WrRd^.astBitStWrRd_Switch_Grp[iGrp].xSwitch_UseFollow_1U_V_UwCut					:= i_pstStSysParam^.astStGrpParam_Save[iGrp].xUseFollow_1U_V_UwCut ;(*裁切套色新方式开关*)
	i_pstStParam_Diamonds_WrRd^.astBitStWrRd_Switch_Grp[iGrp].xSwitch_TypeGetInitDiam						:= i_pstStSysParam^.stStSysParam_Save.xTypeGetInitDiam ;(*收放料初始卷径获取方式*)

	i_pstStParam_Diamonds_WrRd^.astBitStWrRd_Switch_Grp[iGrp].xSwitch_Heating_I				:= i_pstStSysParam^.astStGrpParam_UnSave[iGrp].xBtn_AllHeating_I				;//	: BIT;(*全体加热I当*)
	i_pstStParam_Diamonds_WrRd^.astBitStWrRd_Switch_Grp[iGrp].xSwitch_Heating_II			:= i_pstStSysParam^.astStGrpParam_UnSave[iGrp].xBtn_AllHeating_II		  		;//	: BIT;(*全体加热II当*)
	i_pstStParam_Diamonds_WrRd^.astBitStWrRd_Switch_Grp[iGrp].xSwitch_Heating_III			:= i_pstStSysParam^.astStGrpParam_UnSave[iGrp].xBtn_AllHeating_III				;//    : BIT;(*全体加热III当*)
	i_pstStParam_Diamonds_WrRd^.astBitStWrRd_Switch_Grp[iGrp].xSwitch_Heating_Close			:= i_pstStSysParam^.astStGrpParam_UnSave[iGrp].xBtn_AllHeating_Close			;//	: BIT;(*全体加热关*)
	i_pstStParam_Diamonds_WrRd^.astBitStWrRd_Switch_Grp[iGrp].xSwitch_Heating_Water			:= i_pstStSysParam^.astStGrpParam_UnSave[iGrp].xBtn_AllHeating_Water	 		;//    : BIT;	(*全体水加热*)
	i_pstStParam_Diamonds_WrRd^.astBitStWrRd_Switch_Grp[iGrp].xSwitch_Heating_Elc			:= i_pstStSysParam^.astStGrpParam_UnSave[iGrp].xBtn_AllHeating_Elc				;//	: BIT;(*全体电加热*)
	i_pstStParam_Diamonds_WrRd^.astBitStWrRd_Switch_Grp[iGrp].xBtn_CopySV_1U_To_Other		:= i_pstStSysParam^.astStGrpParam_UnSave[iGrp].xBtn_CopySV_1U_To_Other			;//	: BIT;(*复制1U排风频率到所有色*)
	i_pstStParam_Diamonds_WrRd^.astBitStWrRd_Switch_Grp[iGrp].xBtn_Reset_TempCtlBlock		:= i_pstStSysParam^.astStGrpParam_UnSave[iGrp].xBtn_Reset_TempCtlBlock			;//	: BIT;(*复位温控模块按钮*)
	i_pstStParam_Diamonds_WrRd^.astBitStWrRd_Switch_Grp[iGrp].xBtn_AllExhAir_On				:= i_pstStSysParam^.astStGrpParam_UnSave[iGrp].xBtn_AllExhAir_On				;//	: BIT;(*全体排风开*)
	i_pstStParam_Diamonds_WrRd^.astBitStWrRd_Switch_Grp[iGrp].xBtn_AllExhAir_Off			:= i_pstStSysParam^.astStGrpParam_UnSave[iGrp].xBtn_AllExhAir_Off				;//	: BIT;(*全体排风关*)
	i_pstStParam_Diamonds_WrRd^.astBitStWrRd_Switch_Grp[iGrp].xBtn_CopyExhFreq_1U_To_Other	:= i_pstStSysParam^.astStGrpParam_UnSave[iGrp].xBtn_CopyExhFreq_1U_To_Other	;//	: BIT;(*复制1U排风频率到所有色*)
	i_pstStParam_Diamonds_WrRd^.astBitStWrRd_Switch_Grp[iGrp].xBtn_ExhAir_Reset				:= i_pstStSysParam^.astStGrpParam_UnSave[iGrp].xBtn_ExhAir_Reset				;//	: BIT;(*排风复位按钮*)

	i_pstStParam_Diamonds_WrRd^.astBitStWrRd_Switch_Grp[iGrp].xPidType_If_New								:= i_pstStSysParam^.astStGrpParam_Save[iGrp].xPidType_If_New;
	i_pstStParam_Diamonds_WrRd^.astBitStWrRd_Switch_Grp[iGrp].xPidType_Of_New                 				:= i_pstStSysParam^.astStGrpParam_Save[iGrp].xPidType_Of_New;
	i_pstStParam_Diamonds_WrRd^.astBitStWrRd_Switch_Grp[iGrp].xBtn_StepTest_V                 				:= i_pstStSysParam^.astStGrpParam_UnSave[iGrp].xBtn_StepTest_V;
	i_pstStParam_Diamonds_WrRd^.astBitStWrRd_Switch_Grp[iGrp].xUseDiam_LowPass_Rw             				:= i_pstStSysParam^.astStGrpParam_Save[iGrp].xUseDiam_LowPass_Rw;
	i_pstStParam_Diamonds_WrRd^.astBitStWrRd_Switch_Grp[iGrp].xTensionCompensateEn_Rw         				:= i_pstStSysParam^.astStGrpParam_Save[iGrp].xTensionCompensateEn_Rw;
	i_pstStParam_Diamonds_WrRd^.astBitStWrRd_Switch_Grp[iGrp].xUseTime_b1_Rw                  				:= i_pstStSysParam^.astStGrpParam_Save[iGrp].xUseTime_b1_Rw;
	i_pstStParam_Diamonds_WrRd^.astBitStWrRd_Switch_Grp[iGrp].xUseTime_Variaition_Rw          				:= i_pstStSysParam^.astStGrpParam_Save[iGrp].xUseTime_Variaition_Rw;
	i_pstStParam_Diamonds_WrRd^.astBitStWrRd_Switch_Grp[iGrp].xUseIMatrix_rX_DARE_Rw          				:= i_pstStSysParam^.astStGrpParam_Save[iGrp].xUseIMatrix_rX_DARE_Rw;
	i_pstStParam_Diamonds_WrRd^.astBitStWrRd_Switch_Grp[iGrp].xTensionCompensateEn_RwCut      				:= i_pstStSysParam^.astStGrpParam_Save[iGrp].xTensionCompensateEn_RwCut;
	i_pstStParam_Diamonds_WrRd^.astBitStWrRd_Switch_Grp[iGrp].xUseDiam_LowPass_Uw             				:= i_pstStSysParam^.astStGrpParam_Save[iGrp].xUseDiam_LowPass_Uw;
	i_pstStParam_Diamonds_WrRd^.astBitStWrRd_Switch_Grp[iGrp].xTensionCompensateEn_Uw         				:= i_pstStSysParam^.astStGrpParam_Save[iGrp].xTensionCompensateEn_Uw;
	i_pstStParam_Diamonds_WrRd^.astBitStWrRd_Switch_Grp[iGrp].xUseTime_b1_Uw                  				:= i_pstStSysParam^.astStGrpParam_Save[iGrp].xUseTime_b1_Uw;
	i_pstStParam_Diamonds_WrRd^.astBitStWrRd_Switch_Grp[iGrp].xUseTime_Variaition_Uw          				:= i_pstStSysParam^.astStGrpParam_Save[iGrp].xUseTime_Variaition_Uw;
	i_pstStParam_Diamonds_WrRd^.astBitStWrRd_Switch_Grp[iGrp].xUseIMatrix_rX_DARE_Uw          				:= i_pstStSysParam^.astStGrpParam_Save[iGrp].xUseIMatrix_rX_DARE_Uw;

	i_pstStParam_Diamonds_WrRd^.astBitStWrRd_Switch_Grp[iGrp].xSwitch_Estimate_Uw:= i_pstStSysParam^.astStGrpParam_Save[iGrp].xDiaEstEn_Uw;
	i_pstStParam_Diamonds_WrRd^.astBitStWrRd_Switch_Grp[iGrp].xSwitch_Estimate_Rw:= i_pstStSysParam^.astStGrpParam_Save[iGrp].xDiaEstEn_Rw;

	i_pstStParam_Diamonds_WrRd^.astBitStWrRd_Switch_Grp[iGrp].xSwitchTension_If:= i_pstStSysParam^.astStGrpParam_Save[iGrp].xSwitchTension_If;
	i_pstStParam_Diamonds_WrRd^.astBitStWrRd_Switch_Grp[iGrp].xSwitchTension_Of:= i_pstStSysParam^.astStGrpParam_Save[iGrp].xSwitchTension_Of;
	//2025.9.18.171636
	i_pstStParam_Diamonds_WrRd^.astBitStWrRd_Switch_Grp[iGrp].xNegPolarity_Uw:= i_pstStSysParam^.astStGrpParam_Save[iGrp].wAI_polarity.0;
	i_pstStParam_Diamonds_WrRd^.astBitStWrRd_Switch_Grp[iGrp].xNegPolarity_Rw:= i_pstStSysParam^.astStGrpParam_Save[iGrp].wAI_polarity.1;
	i_pstStParam_Diamonds_WrRd^.astBitStWrRd_Switch_Grp[iGrp].xNegPolarity_If:= i_pstStSysParam^.astStGrpParam_Save[iGrp].wAI_polarity.2;
	i_pstStParam_Diamonds_WrRd^.astBitStWrRd_Switch_Grp[iGrp].xNegPolarity_Of:= i_pstStSysParam^.astStGrpParam_Save[iGrp].wAI_polarity.3;

	i_pstStParam_Diamonds_WrRd^.astBitStWrRd_Switch_Grp[iGrp].xUseBtn_Linkage:= i_pstStSysParam^.astStGrpParam_Save[iGrp].xUseBtn_Linkage;
	i_pstStParam_Diamonds_WrRd^.astBitStWrRd_Switch_Grp[iGrp].xSwitch_ScraperOn_Of:= i_pstStSysParam^.astStGrpParam_Save[iGrp].xSwitch_ScraperOn_Of;
(*2025.10.24.144602*)
	i_pstStParam_Diamonds_WrRd^.astBitStWrRd_Switch_Grp[iGrp].xSwitch_TempFromEnc_PT1000_If:= i_pstStSysParam^.astStGrpParam_Save[iGrp].xSwitch_TempFromEnc_PT1000_If;
	i_pstStParam_Diamonds_WrRd^.astBitStWrRd_Switch_Grp[iGrp].xSwitch_TempFromEnc_PT1000_Of:= i_pstStSysParam^.astStGrpParam_Save[iGrp].xSwitch_TempFromEnc_PT1000_Of;
	i_pstStParam_Diamonds_WrRd^.astBitStWrRd_Switch_Grp[iGrp].xSwitch_MotorTemp_PT1000_NTC_If:= i_pstStSysParam^.astStGrpParam_Save[iGrp].xSwitch_MotorTemp_PT1000_NTC_If;
	i_pstStParam_Diamonds_WrRd^.astBitStWrRd_Switch_Grp[iGrp].xSwitch_MotorTemp_PT1000_NTC_Of:= i_pstStSysParam^.astStGrpParam_Save[iGrp].xSwitch_MotorTemp_PT1000_NTC_Of;
	i_pstStParam_Diamonds_WrRd^.astBitStWrRd_Switch_Grp[iGrp].xTensionCompensateEn_UwCut:= i_pstStSysParam^.astStGrpParam_Save[iGrp].xTensionCompensateEn_UwCut;
	i_pstStParam_Diamonds_WrRd^.astBitStWrRd_Switch_Grp[iGrp].xUseAntiNotch_Uw:= i_pstStSysParam^.astStGrpParam_Save[iGrp].xUseAntiNotch_Uw;
	i_pstStParam_Diamonds_WrRd^.astBitStWrRd_Switch_Grp[iGrp].xWorkMode_RollerPress:= i_pstStSysParam^.astStGrpParam_Save[iGrp].xWorkMode_RollerPress;
	i_pstStParam_Diamonds_WrRd^.astBitStWrRd_Switch_Grp[iGrp].xSwitch_WaitFilmLengthEn:= i_pstStSysParam^.astStGrpParam_Save[iGrp].xSwitch_WaitFilmLengthEn;
	i_pstStParam_Diamonds_WrRd^.astBitStWrRd_Switch_Grp[iGrp].xSwitch_WaitFilmLengthEn_From1st:= i_pstStSysParam^.astStGrpParam_Save[iGrp].xSwitch_WaitFilmLengthEn_From1st;
	i_pstStParam_Diamonds_WrRd^.astBitStWrRd_Switch_Grp[iGrp].xSwitch_Alarm_Arc:= i_pstStSysParam^.astStGrpParam_Save[iGrp].xSwitch_Alarm_Arc;
	i_pstStParam_Diamonds_WrRd^.astBitStWrRd_Switch_Grp[iGrp].xSwitch_PreHotAirEn:= i_pstStSysParam^.astStGrpParam_Save[iGrp].xSwitch_PreHotAirEn;
	i_pstStParam_Diamonds_WrRd^.astBitStWrRd_Switch_Grp[iGrp].xSwitch_PreHeatingEn:= i_pstStSysParam^.astStGrpParam_Save[iGrp].xSwitch_PreHeatingEn;

	i_pstStParam_Diamonds_WrRd^.astBitStWrRd_Switch_Grp[iGrp].xBtn_PreRegisterAxisId_Manu:= i_pstStSysParam^.astStGrpParam_UnSave[iGrp].xBtn_PreRegisterAxisId_Manu;
	i_pstStParam_Diamonds_WrRd^.astBitStWrRd_Switch_Grp[iGrp].xBtn_PreRegister:= i_pstStSysParam^.astStGrpParam_UnSave[iGrp].xBtn_PreRegister;
	i_pstStParam_Diamonds_WrRd^.astBitStWrRd_Switch_Grp[iGrp].xBtn_PreRegisterCorrConfirm:= i_pstStSysParam^.astStGrpParam_UnSave[iGrp].xBtn_PreRegisterCorrConfirm;
	i_pstStParam_Diamonds_WrRd^.astBitStWrRd_Switch_Grp[iGrp].xBtn_HorzPreRegister_Repeat:= i_pstStSysParam^.astStGrpParam_UnSave[iGrp].xBtn_HorzPreRegister_Repeat;
	i_pstStParam_Diamonds_WrRd^.astBitStWrRd_Switch_Grp[iGrp].xBtn_HorzPreRegister_Setup:= i_pstStSysParam^.astStGrpParam_UnSave[iGrp].xBtn_HorzPreRegister_Setup;

	(*待补充-结束|2025.08.06.215042*)
	i_pstStParam_Diamonds_WrRd^.adwDiamAlarm_Uw[iGrp]														:= REAL_TO_DWORD(i_pstStSysParam^.astStGrpParam_Save[iGrp].rDiamAlarm_Uw);				(*放料报警卷径*)
	i_pstStParam_Diamonds_WrRd^.arFilmThickNess_Using[iGrp]													:= i_pstStSysParam^.astStGrpParam_Save[iGrp].rFilmThickNess_Using;						(*料膜厚度手动输入值*)
	i_pstStParam_Diamonds_WrRd^.arInitTaper_Hmi_Rw[iGrp]													:= i_pstStSysParam^.astStGrpParam_Save[iGrp].rInitTaper_Hmi_Rw;							(*收料起始气压*)
	i_pstStParam_Diamonds_WrRd^.auiVel_CommonlyUsed[iGrp,1]												:= REAL_TO_UINT(i_pstStSysParam^.astStGrpParam_Save[iGrp].arVel_Usr[1]);						(*常用速度*)
	i_pstStParam_Diamonds_WrRd^.auiVel_CommonlyUsed[iGrp,2]												:= REAL_TO_UINT(i_pstStSysParam^.astStGrpParam_Save[iGrp].arVel_Usr[2]);						(*常用速度*)
	i_pstStParam_Diamonds_WrRd^.auiVel_CommonlyUsed[iGrp,3]												:= REAL_TO_UINT(i_pstStSysParam^.astStGrpParam_Save[iGrp].arVel_Usr[3]);						(*常用速度*)
	i_pstStParam_Diamonds_WrRd^.aiCutDneResetPidMultiple_Uw[iGrp]											:= i_pstStSysParam^.astStGrpParam_Save[iGrp].iCutDneResetPidMultiple_Uw;				(*裁切PID放大系数-放料*)
	i_pstStParam_Diamonds_WrRd^.aiCutDneResetPidRemainTime_Uw[iGrp]											:= i_pstStSysParam^.astStGrpParam_Save[iGrp].iCutDneResetPidRemainTime_Uw;				(*裁切PID放大保持时间-放料*)
	i_pstStParam_Diamonds_WrRd^.aiCutDneResetPidDefaultTime_Uw[iGrp]										:= i_pstStSysParam^.astStGrpParam_Save[iGrp].iCutDneResetPidToDefaultTime_Uw;			(*裁切PID放大恢复时间-放料*)
	i_pstStParam_Diamonds_WrRd^.aiCutDneResetPidMultiple_Rw[iGrp]											:= i_pstStSysParam^.astStGrpParam_Save[iGrp].iCutDneResetPidMultiple_Rw;				(*裁切PID放大系数-收料*)
	i_pstStParam_Diamonds_WrRd^.aiCutDneResetPidRemainTime_Rw[iGrp]											:= i_pstStSysParam^.astStGrpParam_Save[iGrp].iCutDneResetPidRemainTime_Rw;				(*裁切PID放大保持时间-收料*)
	i_pstStParam_Diamonds_WrRd^.aiCutDneResetPidDefaultTime_Rw[iGrp]										:= i_pstStSysParam^.astStGrpParam_Save[iGrp].iCutDneResetPidToDefaultTime_Rw;			(*裁切PID放大恢复时间-收料*)
	i_pstStParam_Diamonds_WrRd^.abyAutoMaticCutMode_uw[iGrp]												:= i_pstStSysParam^.astStGrpParam_Save[iGrp].byAutoMaticCutMode_uw;						(*放料自动接料方式-剩余卷径/剩余米数*)

	i_pstStParam_Diamonds_WrRd^.arDia_PaperRoller_Uw[iGrp]			:= i_pstStSysParam^.astStGrpParam_Save[iGrp].rDia_PaperRoller_Uw;							(*放料纸筒直径*)
	i_pstStParam_Diamonds_WrRd^.auiAutoMaticCutDia_Uw[iGrp]			:= i_pstStSysParam^.astStGrpParam_Save[iGrp].uiAutoMaticCutDia_Uw;							(*放料剩余卷径*)
	i_pstStParam_Diamonds_WrRd^.auiAutoMaticCutMeters_Uw[iGrp]		:= i_pstStSysParam^.astStGrpParam_Save[iGrp].uiAutoMaticCutMeters_Uw;						(*放料剩余米数*)
	i_pstStParam_Diamonds_WrRd^.abyAutoMaticCutMode_Rw[iGrp]		:= i_pstStSysParam^.astStGrpParam_Save[iGrp].byAutoMaticCutMode_Rw;							(*收料自动接料方式-收料米数/整机料长*)
	i_pstStParam_Diamonds_WrRd^.auiAutoMaticCutMeters_Rw[iGrp]		:= i_pstStSysParam^.astStGrpParam_Save[iGrp].uiAutoMaticCutMeters_Rw;						(*收料米数*)
	i_pstStParam_Diamonds_WrRd^.abyLenth_Machine[iGrp]				:= i_pstStSysParam^.astStGrpParam_Save[iGrp].byLenth_Machine;								(*整机料长*)
	i_pstStParam_Diamonds_WrRd^.arPressure_Max[iGrp]				:= i_pstStSysParam^.astStGrpParam_Save[iGrp].rPressure_Max;									(*涂布压力传感器最大标定压力值*)
	i_pstStParam_Diamonds_WrRd^.arHz_MainExhaust_ManuallySet[iGrp]	:= i_pstStSysParam^.astStGrpParam_Save[iGrp].rHz_MainExhaust_ManuallySet;					(*主排风手动频率*)
	i_pstStParam_Diamonds_WrRd^.aiMarkId[iGrp]						:= i_pstStSysParam^.astStGrpParam_Save[iGrp].iMarkTypeId;									(*色斑形式*)
	i_pstStParam_Diamonds_WrRd^.aicurMarkArrangeId[iGrp]			:= i_pstStSysParam^.astStGrpParam_Save[iGrp].iMarkArrangeMode;								(*色标顺序*)
	i_pstStParam_Diamonds_WrRd^.abyTriMark_SideC[iGrp]				:= i_pstStSysParam^.astStGrpParam_Save[iGrp].byTriMark_SideC;								(*梯标直边宽度1mm*)
	i_pstStParam_Diamonds_WrRd^.abyTriMark_SideB[iGrp]				:= i_pstStSysParam^.astStGrpParam_Save[iGrp].byTriMark_SideB;								(*梯标直边宽度2mm*)
	i_pstStParam_Diamonds_WrRd^.arAI_med_Uw[iGrp]					:= i_pstStSysParam^.astStGrpParam_Save[iGrp].rAI_med_Uw;									(*放料摆臂中位值/rAI_med_Uw*)
	i_pstStParam_Diamonds_WrRd^.arAI_med_Rw[iGrp]					:= i_pstStSysParam^.astStGrpParam_Save[iGrp].rAI_med_Rw;									(*收料摆臂中位值/rAI_med_Rw*)
	i_pstStParam_Diamonds_WrRd^.arAI_med_If[iGrp]					:= i_pstStSysParam^.astStGrpParam_Save[iGrp].rAI_med_If;									(*放牵摆臂中位值/rAI_med_If*)
	i_pstStParam_Diamonds_WrRd^.arAI_med_Of[iGrp]					:= i_pstStSysParam^.astStGrpParam_Save[iGrp].rAI_med_Of;									(*收牵摆臂中位值/rAI_med_Of*)
	i_pstStParam_Diamonds_WrRd^.arRatedRpm_Uw[iGrp]					:= INT_TO_REAL(i_pstStSysParam^.astStGrpParam_Save[iGrp].iRatedRpm_Uw);						(*额定转速*)
	i_pstStParam_Diamonds_WrRd^.arRatedFreq_Uw[iGrp]				:= INT_TO_REAL(i_pstStSysParam^.astStGrpParam_Save[iGrp].iRatedFreq_Uw);					(*额定频率*)
	i_pstStParam_Diamonds_WrRd^.arUpperFreq_Uw[iGrp]				:= INT_TO_REAL(i_pstStSysParam^.astStGrpParam_Save[iGrp].iUpperFreq_Uw);					(*上限频率*)
	i_pstStParam_Diamonds_WrRd^.arRatedRpm_Rw[iGrp]					:= INT_TO_REAL(i_pstStSysParam^.astStGrpParam_Save[iGrp].iRatedRpm_Rw);						(*额定转速*)
	i_pstStParam_Diamonds_WrRd^.arRatedFreq_Rw[iGrp]				:= INT_TO_REAL(i_pstStSysParam^.astStGrpParam_Save[iGrp].iRatedFreq_Rw);					(*额定频率*)
	i_pstStParam_Diamonds_WrRd^.arUpperFreq_Rw[iGrp]				:= INT_TO_REAL(i_pstStSysParam^.astStGrpParam_Save[iGrp].iUpperFreq_Rw);					(*上限频率*)
	i_pstStParam_Diamonds_WrRd^.arRatedRpm_If[iGrp]					:= INT_TO_REAL(i_pstStSysParam^.astStGrpParam_Save[iGrp].iRatedRpm_If);						(*额定转速*)
	i_pstStParam_Diamonds_WrRd^.arRatedFreq_If[iGrp]				:= INT_TO_REAL(i_pstStSysParam^.astStGrpParam_Save[iGrp].iRatedFreq_If);					(*额定频率*)
	i_pstStParam_Diamonds_WrRd^.arUpperFreq_If[iGrp]				:= INT_TO_REAL(i_pstStSysParam^.astStGrpParam_Save[iGrp].iUpperFreq_If);					(*上限频率*)
	i_pstStParam_Diamonds_WrRd^.arRatedRpm_Of[iGrp]					:= INT_TO_REAL(i_pstStSysParam^.astStGrpParam_Save[iGrp].iRatedRpm_Of);						(*额定转速*)
	i_pstStParam_Diamonds_WrRd^.arRatedFreq_Of[iGrp]				:= INT_TO_REAL(i_pstStSysParam^.astStGrpParam_Save[iGrp].iRatedFreq_Of);					(*额定频率*)
	i_pstStParam_Diamonds_WrRd^.arUpperFreq_Of[iGrp]				:= INT_TO_REAL(i_pstStSysParam^.astStGrpParam_Save[iGrp].iUpperFreq_Of);					(*上限频率*)
	i_pstStParam_Diamonds_WrRd^.arDiamTaper_Begin_Rw[iGrp]			:= i_pstStSysParam^.astStGrpParam_Save[iGrp].rDiam_taper_begin_Rw;							(*锥度起始直径*)
	i_pstStParam_Diamonds_WrRd^.arDiamTaper_End_Rw[iGrp]            := i_pstStSysParam^.astStGrpParam_Save[iGrp].rDiam_taper_end_Rw;							(*锥度结束直径*)
	i_pstStParam_Diamonds_WrRd^.arGirth_3Inch[iGrp]                 := i_pstStSysParam^.astStGrpParam_Save[iGrp].rGirth_3inch_Rw;								(*收料3吋默认周长*)
	i_pstStParam_Diamonds_WrRd^.arGirth_6Inch[iGrp]                 := i_pstStSysParam^.astStGrpParam_Save[iGrp].rGirth_6inch_Rw;								(*收料6吋默认周长*)
	i_pstStParam_Diamonds_WrRd^.abyAIType_Uw[iGrp]:= i_pstStSysParam^.astStGrpParam_Save[iGrp].byAIType_Uw;
	i_pstStParam_Diamonds_WrRd^.abyAIType_Rw[iGrp]:= i_pstStSysParam^.astStGrpParam_Save[iGrp].byAIType_Rw;
	i_pstStParam_Diamonds_WrRd^.abyAIType_If[iGrp]:= i_pstStSysParam^.astStGrpParam_Save[iGrp].byAIType_If;
	i_pstStParam_Diamonds_WrRd^.abyAIType_Of[iGrp]:= i_pstStSysParam^.astStGrpParam_Save[iGrp].byAIType_Of;

	i_pstStParam_Diamonds_WrRd^.arKpid_SVol_Uw[iGrp,1]	  := i_pstStSysParam^.astStGrpParam_Save[iGrp].arKpid_Uw[1];											(*放料PID设定*)
	i_pstStParam_Diamonds_WrRd^.arKpid_SVol_Uw[iGrp,2]	  := i_pstStSysParam^.astStGrpParam_Save[iGrp].arKpid_Uw[2];											(*放料PID设定*)
	i_pstStParam_Diamonds_WrRd^.arKpid_SVol_Uw[iGrp,3]	  := i_pstStSysParam^.astStGrpParam_Save[iGrp].arKpid_Uw[3];											(*放料PID设定*)

	i_pstStParam_Diamonds_WrRd^.arKpid_SVol_Rw[iGrp,1]	  := i_pstStSysParam^.astStGrpParam_Save[iGrp].arKpid_Rw[1];											(*收料PID设定*)
	i_pstStParam_Diamonds_WrRd^.arKpid_SVol_Rw[iGrp,2]	  := i_pstStSysParam^.astStGrpParam_Save[iGrp].arKpid_Rw[2];											(*收料PID设定*)
	i_pstStParam_Diamonds_WrRd^.arKpid_SVol_Rw[iGrp,3]	  := i_pstStSysParam^.astStGrpParam_Save[iGrp].arKpid_Rw[3];											(*收料PID设定*)

	i_pstStParam_Diamonds_WrRd^.arKpid_If[iGrp,1]			  := i_pstStSysParam^.astStGrpParam_Save[iGrp].arKpid_If[1];											(*放牵PID设定*)
	i_pstStParam_Diamonds_WrRd^.arKpid_If[iGrp,2]			  := i_pstStSysParam^.astStGrpParam_Save[iGrp].arKpid_If[2];											(*放牵PID设定*)
	i_pstStParam_Diamonds_WrRd^.arKpid_If[iGrp,3]			  := i_pstStSysParam^.astStGrpParam_Save[iGrp].arKpid_If[3];											(*放牵PID设定*)

	i_pstStParam_Diamonds_WrRd^.arKpid_Of[iGrp,1]			  := i_pstStSysParam^.astStGrpParam_Save[iGrp].arKpid_Of[1];											(*收牵PID设定*)
	i_pstStParam_Diamonds_WrRd^.arKpid_Of[iGrp,2]			  := i_pstStSysParam^.astStGrpParam_Save[iGrp].arKpid_Of[2];											(*收牵PID设定*)
	i_pstStParam_Diamonds_WrRd^.arKpid_Of[iGrp,3]			  := i_pstStSysParam^.astStGrpParam_Save[iGrp].arKpid_Of[3];											(*收牵PID设定*)

	i_pstStParam_Diamonds_WrRd^.abyCoef_Stiffen_Uw[iGrp]                      := i_pstStSysParam^.astStGrpParam_Save[iGrp].byCoef_Stiffen_Uw;						(*放料拉料系数*)
	i_pstStParam_Diamonds_WrRd^.abyCoef_Stiffen_Rw[iGrp]                      := i_pstStSysParam^.astStGrpParam_Save[iGrp].byCoef_Stiffen_Rw;						(*收料拉料系数*)
	i_pstStParam_Diamonds_WrRd^.abyInitialSpd_Stiffen[iGrp]                   := i_pstStSysParam^.astStGrpParam_Save[iGrp].byInitialSpd_Stiffen_Uw;					(*拉料初始速度*)
	i_pstStParam_Diamonds_WrRd^.abyStationIdDst_VirEnc[iGrp]                  := i_pstStSysParam^.astStGrpParam_Save[iGrp].byStationIdDst_VirEnc;					(*异站编码器目标站好*)
	i_pstStParam_Diamonds_WrRd^.abyDelayTime_DiaCompensateWhenCutDne_Uw[iGrp] := i_pstStSysParam^.astStGrpParam_Save[iGrp].byDelayTime_DiaCompensateWhenCutDne_Uw;  (*放料裁切延时*)
	i_pstStParam_Diamonds_WrRd^.abyVelSa_DiamCompensate_Uw[iGrp]			  := i_pstStSysParam^.astStGrpParam_Save[iGrp].byVelSa_DiamCompensate_Uw;				(*放料补偿速度*)
	i_pstStParam_Diamonds_WrRd^.abyDelayTime_DiaCompensateWhenCutDne_Rw[iGrp] := i_pstStSysParam^.astStGrpParam_Save[iGrp].byDelayTime_DiaCompensateWhenCutDne_Rw;	(*收料裁切延时*)
	i_pstStParam_Diamonds_WrRd^.abyVelSa_DiamCompensate_Rw[iGrp]			  := i_pstStSysParam^.astStGrpParam_Save[iGrp].byVelSa_DiamCompensate_Rw;				(*收料补偿速度*)
	i_pstStParam_Diamonds_WrRd^.arRatedRpm_Scraper[iGrp]					  := LREAL_TO_REAL(i_pstStSysParam^.astStGrpParam_Save[iGrp].lrRatedRpm_Scraper);		(*刮刀额定转速*)
	i_pstStParam_Diamonds_WrRd^.arRatedFreq_Scraper[iGrp]	                  := LREAL_TO_REAL(i_pstStSysParam^.astStGrpParam_Save[iGrp].lrRatedFreq_Scraper);		(*刮刀额定频率*)
	i_pstStParam_Diamonds_WrRd^.arUpperFreq_Scraper[iGrp]                 	  := LREAL_TO_REAL(i_pstStSysParam^.astStGrpParam_Save[iGrp].lrUpperFreq_Scraper);		(*刮刀上限频率*)
	i_pstStParam_Diamonds_WrRd^.arMinFreq_Scraper[iGrp]                   	  := (i_pstStSysParam^.astStGrpParam_Save[iGrp].rMinFreq_Scraper);		(*刮刀最小频率*)
	i_pstStParam_Diamonds_WrRd^.arMaxFreq_Scraper[iGrp]                   	  := (i_pstStSysParam^.astStGrpParam_Save[iGrp].rMaxFreq_Scraper);		(*刮刀最大频率*)
	i_pstStParam_Diamonds_WrRd^.aiRatio_ScraperContrastToPrintRoller[iGrp]	  := i_pstStSysParam^.astStGrpParam_Save[iGrp].iRatio_ScraperContrastToPrintRoller;		(*刮刀调整比例*)
	i_pstStParam_Diamonds_WrRd^.aiVelSa_ScraperRun[iGrp]                  	  := i_pstStSysParam^.astStGrpParam_Save[iGrp].iVelSa_ScraperRun;						(*刮刀启动速度*)
	i_pstStParam_Diamonds_WrRd^.aiDen_ScraperMotor[iGrp]                  	  := i_pstStSysParam^.astStGrpParam_Save[iGrp].iDen_ScraperMotor;						(*刮刀减速比分母*)
	i_pstStParam_Diamonds_WrRd^.aiNum_ScraperMotor[iGrp]                  	  := i_pstStSysParam^.astStGrpParam_Save[iGrp].iNum_ScraperMotor;						(*刮刀减速比分子*)
	i_pstStParam_Diamonds_WrRd^.aiUpperFreq_InkRoller[iGrp]               	  := i_pstStSysParam^.astStGrpParam_Save[iGrp].iUpperFreq_InkRoller;					(*递磨辊上限频率*)
	i_pstStParam_Diamonds_WrRd^.aiVelSa_InkRollerRun[iGrp]                	  := i_pstStSysParam^.astStGrpParam_Save[iGrp].iVelSa_InkRollerRun;						(*递磨辊启动速度*)
	i_pstStParam_Diamonds_WrRd^.aiFrq_InkRollerMin[iGrp]                  	  := i_pstStSysParam^.astStGrpParam_Save[iGrp].iFrq_InkRollerMin;						(*递磨辊最小频率*)
	i_pstStParam_Diamonds_WrRd^.aiFrq_InkRollerMax[iGrp]                  	  := i_pstStSysParam^.astStGrpParam_Save[iGrp].iFrq_InkRollerMax;						(*递磨辊最大频率*)
	i_pstStParam_Diamonds_WrRd^.aiVel_InkRollerMin[iGrp]                  	  := i_pstStSysParam^.astStGrpParam_Save[iGrp].iVel_InkRollerMin;						(*递磨辊最小速度*)
	i_pstStParam_Diamonds_WrRd^.aiVel_InkRollerMax[iGrp]                  	  := i_pstStSysParam^.astStGrpParam_Save[iGrp].iVel_InkRollerMax;						(*递磨辊最大速度*)
	i_pstStParam_Diamonds_WrRd^.abyPseudoRandomId[iGrp]:=	i_pstStSysParam^.astStGrpParam_UnSave[iGrp].byPseudoRandomId;
	i_pstStParam_Diamonds_WrRd^.abyFilmType[iGrp]:= i_pstStSysParam^.astStGrpParam_Save[iGrp].byFilmType;
	i_pstStParam_Diamonds_WrRd^.auiUseTime_Diam_Min_Uw[iGrp]:= i_pstStSysParam^.astStGrpParam_Save[iGrp].uiUseTime_Diam_Min_Uw;
	i_pstStParam_Diamonds_WrRd^.auiUseTime_Diam_Min_Rw[iGrp]:= i_pstStSysParam^.astStGrpParam_Save[iGrp].uiUseTime_Diam_Min_Rw;

	i_pstStParam_Diamonds_WrRd^.aiPreHotRoller_Velocity_PreHot[iGrp]   := i_pstStSysParam^.astStGrpParam_Save[iGrp].iPreHotRoller_Velocity_PreHot;  				(*预热辊额定转速*)
	i_pstStParam_Diamonds_WrRd^.arStandardFreq_HotRoller_PreHot[iGrp]  := i_pstStSysParam^.astStGrpParam_Save[iGrp].rStandardFreq_HotRoller_PreHot; 				(*预热辊额定频率*)
	i_pstStParam_Diamonds_WrRd^.arUpperFreq_HotRoller_PreHot[iGrp]     := i_pstStSysParam^.astStGrpParam_Save[iGrp].rUpperFreq_HotRoller_PreHot;    				(*预热辊上限频率*)
	i_pstStParam_Diamonds_WrRd^.arCoeff_HotRoller_PreHot[iGrp]         := i_pstStSysParam^.astStGrpParam_Save[iGrp].rCoeff_HotRoller_PreHot;        				(*预热辊速度系数*)
	i_pstStParam_Diamonds_WrRd^.arGirth_HotRoller_PreHot[iGrp]         := i_pstStSysParam^.astStGrpParam_Save[iGrp].rGirth_HotRoller_PreHot;        				(*预热辊周长*)
	i_pstStParam_Diamonds_WrRd^.aiPreAirHotRollTorque[iGrp]            := i_pstStSysParam^.astStGrpParam_Save[iGrp].iPreAirHotRollTorque;           				(*预热辊转矩*)
	i_pstStParam_Diamonds_WrRd^.auiDen_HotRoller_PreHot[iGrp]          := i_pstStSysParam^.astStGrpParam_Save[iGrp].uiDen_HotRoller_PreHot;         				(*预热辊减速比分母*)
	i_pstStParam_Diamonds_WrRd^.auiNum_HotRoller_PreHot[iGrp]          := i_pstStSysParam^.astStGrpParam_Save[iGrp].uiNum_HotRoller_PreHot;         				(*预热辊减速比分子*)
	i_pstStParam_Diamonds_WrRd^.aiPreHotRoller_Velocity_Water[iGrp]    := i_pstStSysParam^.astStGrpParam_Save[iGrp].iPreHotRoller_Velocity_Water;   				(*水冷辊额定转速*)
	i_pstStParam_Diamonds_WrRd^.arStandardFreq_HotRoller_Water[iGrp]   := i_pstStSysParam^.astStGrpParam_Save[iGrp].rStandardFreq_HotRoller_Water;  				(*水冷辊额定频率*)
	i_pstStParam_Diamonds_WrRd^.arUpperFreq_HotRoller_Water[iGrp]      := i_pstStSysParam^.astStGrpParam_Save[iGrp].rUpperFreq_HotRoller_Water;     				(*水冷辊上限频率*)
	i_pstStParam_Diamonds_WrRd^.arCoeff_HotRoller_Water[iGrp]          := i_pstStSysParam^.astStGrpParam_Save[iGrp].rCoeff_HotRoller_Water;         				(*水冷辊速度系数*)
	i_pstStParam_Diamonds_WrRd^.arGirth_HotRoller_Water[iGrp]          := i_pstStSysParam^.astStGrpParam_Save[iGrp].rGirth_HotRoller_Water;         				(*水冷辊周长*)
	i_pstStParam_Diamonds_WrRd^.auiDen_HotRoller_Water[iGrp]           := i_pstStSysParam^.astStGrpParam_Save[iGrp].uiDen_HotRoller_Water;          				(*水冷辊减速比分母*)
	i_pstStParam_Diamonds_WrRd^.auiNum_HotRoller_Water[iGrp]			:= i_pstStSysParam^.astStGrpParam_Save[iGrp].uiNum_HotRoller_Water;							(*水冷辊减速比分子*)
	i_pstStParam_Diamonds_WrRd^.aiDelayMsec_ExhPowerMode[iGrp]		 	:= i_pstStSysParam^.astStGrpParam_Save[iGrp].iDelayMsec_ExhPowerMode;						(*排风切换延时*)
	i_pstStParam_Diamonds_WrRd^.aiDelayMsec_HeatBlower[iGrp]			:= i_pstStSysParam^.astStGrpParam_Save[iGrp].iDelayMsec_HeatBlower;							(*热风延时*)
	i_pstStParam_Diamonds_WrRd^.aiDelayMsec_Heat[iGrp]				 	:= i_pstStSysParam^.astStGrpParam_Save[iGrp].iDelayMsec_Heat;								(*加热延时*)
	i_pstStParam_Diamonds_WrRd^.abyHotBlowerStopDelayTime[iGrp]		 	:= i_pstStSysParam^.astStGrpParam_Save[iGrp].byHotBlowerStopDelayTime;						(*热风停止延时*)
	i_pstStParam_Diamonds_WrRd^.abyFreqMin_HotWind[iGrp]				:= i_pstStSysParam^.astStGrpParam_Save[iGrp].byFreqMin_HotWind;								(*热风最小频率*)
	i_pstStParam_Diamonds_WrRd^.abyFreqMax_HotWind[iGrp]				:= i_pstStSysParam^.astStGrpParam_Save[iGrp].byFreqMax_HotWind;								(*热风最大频率*)
	i_pstStParam_Diamonds_WrRd^.arStdVol_Diam_Axis_Hmi[iGrp,1]			:= LREAL_TO_REAL(i_pstStSysParam^.astStGrpParam_Save[iGrp].astStStdVolParam_DnCut_UpCut[0].alrStdVol_Diam[1]);			(* 标准卷径值| 双向通讯参数*)
	i_pstStParam_Diamonds_WrRd^.arStdVol_Diam_Axis_Hmi[iGrp,2]			:= LREAL_TO_REAL(i_pstStSysParam^.astStGrpParam_Save[iGrp].astStStdVolParam_DnCut_UpCut[0].alrStdVol_Diam[2]);			(* 标准卷径值| 双向通讯参数*)
	i_pstStParam_Diamonds_WrRd^.arStdVol_Diam_Axis_Hmi[iGrp,3]			:= LREAL_TO_REAL(i_pstStSysParam^.astStGrpParam_Save[iGrp].astStStdVolParam_DnCut_UpCut[0].alrStdVol_Diam[3]);			(* 标准卷径值| 双向通讯参数*)
	i_pstStParam_Diamonds_WrRd^.arStdVol_Diam_Axis_Hmi[iGrp,4]			:= LREAL_TO_REAL(i_pstStSysParam^.astStGrpParam_Save[iGrp].astStStdVolParam_DnCut_UpCut[0].alrStdVol_Diam[4]);			(* 标准卷径值| 双向通讯参数*)
	i_pstStParam_Diamonds_WrRd^.arStdVol_Diam_Axis_Hmi[iGrp,1]			:= LREAL_TO_REAL(i_pstStSysParam^.astStGrpParam_Save[iGrp].astStStdVolParam_DnCut_UpCut[1].alrStdVol_Diam[1]);			(* 标准卷径值| 双向通讯参数*)
	i_pstStParam_Diamonds_WrRd^.arStdVol_Diam_Axis_Hmi[iGrp,2]			:= LREAL_TO_REAL(i_pstStSysParam^.astStGrpParam_Save[iGrp].astStStdVolParam_DnCut_UpCut[1].alrStdVol_Diam[2]);			(* 标准卷径值| 双向通讯参数*)
	i_pstStParam_Diamonds_WrRd^.arStdVol_Diam_Axis_Hmi[iGrp,3]			:= LREAL_TO_REAL(i_pstStSysParam^.astStGrpParam_Save[iGrp].astStStdVolParam_DnCut_UpCut[1].alrStdVol_Diam[3]);			(* 标准卷径值| 双向通讯参数*)
	i_pstStParam_Diamonds_WrRd^.arStdVol_Diam_Axis_Hmi[iGrp,4]			:= LREAL_TO_REAL(i_pstStSysParam^.astStGrpParam_Save[iGrp].astStStdVolParam_DnCut_UpCut[1].alrStdVol_Diam[4]);			(* 标准卷径值| 双向通讯参数*)
	(*待补充-开始|2025.08.07.162226*)
// 	i_pstStParam_Diamonds_WrRd^.arStdVol_Coef[iGrp,1]					:= LREAL_TO_REAL(i_pstStSysParam^.astStGrpParam_UnSave[iGrp].alrStdVol_Coef_Axis_Hmi[1]);					 						 (* 标准卷径系数| 双向通讯参数*)
// 	i_pstStParam_Diamonds_WrRd^.arStdVol_Coef[iGrp,2]					:= LREAL_TO_REAL(i_pstStSysParam^.astStGrpParam_UnSave[iGrp].alrStdVol_Coef_Axis_Hmi[2]);					 						 (* 标准卷径系数| 双向通讯参数*)
// 	i_pstStParam_Diamonds_WrRd^.arStdVol_Coef[iGrp,3]					:= LREAL_TO_REAL(i_pstStSysParam^.astStGrpParam_UnSave[iGrp].alrStdVol_Coef_Axis_Hmi[3]);					 						 (* 标准卷径系数| 双向通讯参数*)
	(*待补充-结束|2025.08.07.162244*)
    i_pstStParam_Diamonds_WrRd^.aiTime_FilmAcc[iGrp]					:= i_pstStSysParam^.astStGrpParam_Save[iGrp].iTime_FilmAcc;												(*预驱料膜加速时间*)
    i_pstStParam_Diamonds_WrRd^.aiTime_FilmDec[iGrp]              	 := i_pstStSysParam^.astStGrpParam_Save[iGrp].iTime_FilmDec;              								  	(*预驱料膜减速时间*)
    i_pstStParam_Diamonds_WrRd^.aiTime_PreDrvAcc_Rw[iGrp]         	 := i_pstStSysParam^.astStGrpParam_Save[iGrp].iTime_PreDrvAcc_Rw;         								  	(*收料预驱加速时间*)
    i_pstStParam_Diamonds_WrRd^.aiTime_PreDrvDec_Rw[iGrp]         	 := i_pstStSysParam^.astStGrpParam_Save[iGrp].iTime_PreDrvDec_Rw;         								  	(*收料预驱减速时间*)
    i_pstStParam_Diamonds_WrRd^.aiTime_PreDrvAcc_Uw[iGrp]         	 := i_pstStSysParam^.astStGrpParam_Save[iGrp].iTime_PreDrvAcc_Uw;         								  	(*放料预驱加速时间*)
    i_pstStParam_Diamonds_WrRd^.aiTime_PreDrvDec_Uw[iGrp]         	 := i_pstStSysParam^.astStGrpParam_Save[iGrp].iTime_PreDrvDec_Uw;         								  	(*放料预驱减速时间*)
    i_pstStParam_Diamonds_WrRd^.arFilmLen_NotAdjFront[iGrp]			 := i_pstStSysParam^.astStGrpParam_Save[iGrp].rFilmLen_NotAdjFront;										  	(*料前幅数*)
    i_pstStParam_Diamonds_WrRd^.arFilmLen_NotAdjBack[iGrp]        	 := i_pstStSysParam^.astStGrpParam_Save[iGrp].rFilmLen_NotAdjBack;        								  	(*料后幅数*)
    i_pstStParam_Diamonds_WrRd^.arFilmLen_UnwindToPU1[iGrp]       	 := i_pstStSysParam^.astStGrpParam_Save[iGrp].rFilmLen_UnwindToPU1;       								   	(*裁点到1色距离*)

	i_pstStParam_Diamonds_WrRd^.auiPiDelay_Uw[iGrp]               		 	:= i_pstStSysParam^.astStGrpParam_Save[iGrp].uiPiDelay_Uw;  										(*放料接料PI投入时间*)
	i_pstStParam_Diamonds_WrRd^.aiPreRevLenth_MM_Cutted[iGrp]     		 	:= i_pstStSysParam^.astStGrpParam_Save[iGrp].iPreRevLenth_MM_Cutted_Uw; 							(*裁切反转距离*)
	i_pstStParam_Diamonds_WrRd^.aiPreRevVel_RPM_Cutted[iGrp]      		 	:= i_pstStSysParam^.astStGrpParam_Save[iGrp].iPreRevVel_RPM_Cutted_Uw;    							(*裁切反转速度*)
	i_pstStParam_Diamonds_WrRd^.arCoefCut_FilmVolPerimeter_Uw[iGrp]		 	:= i_pstStSysParam^.astStGrpParam_Save[iGrp].rCoefCut_FilmVolPerimeter_Uw;       				 	(*放料裁切圈数*)
	i_pstStParam_Diamonds_WrRd^.arCoefCut_FilmVolPerimeter_Rw[iGrp]		 	:= i_pstStSysParam^.astStGrpParam_Save[iGrp].rCoefCut_FilmVolPerimeter_Rw;       				 	(*收料裁切圈数*)
	i_pstStParam_Diamonds_WrRd^.arDiam_Tower_Uw[iGrp]					 	:= i_pstStSysParam^.astStGrpParam_Save[iGrp].rDiam_Tower_Uw;           								(*反转架直径*)
	i_pstStParam_Diamonds_WrRd^.arDiam_NextRoller_Uw[iGrp]            	 	:= i_pstStSysParam^.astStGrpParam_Save[iGrp].rDiam_NextRoller_Uw;      								(*下个辊直径*)
	i_pstStParam_Diamonds_WrRd^.arXPos_NextRoller_Uw[iGrp]            	 	:= i_pstStSysParam^.astStGrpParam_Save[iGrp].rXPos_NextRoller_Uw;      								(*下个辊X*)
	i_pstStParam_Diamonds_WrRd^.arYPos_NextRoller_Uw[iGrp]            	 	:= i_pstStSysParam^.astStGrpParam_Save[iGrp].rYPos_NextRoller_Uw;   								(*下个辊Y*)
	i_pstStParam_Diamonds_WrRd^.arDiam_DeflectorRoller_Uw[iGrp]       	 	:= i_pstStSysParam^.astStGrpParam_Save[iGrp].rDiam_DeflectorRoller_Uw; 								(*导向辊直径*)
	i_pstStParam_Diamonds_WrRd^.arDiam_DeflectorRollPos_Uw[iGrp]      	 	:= i_pstStSysParam^.astStGrpParam_Save[iGrp].rDiam_DeflectorRollPos_Uw;								(*AB导向辊长度*)
	i_pstStParam_Diamonds_WrRd^.aiDebugVelmpm_AxisA_Uw[iGrp]			 	:= i_pstStSysParam^.astStGrpParam_UnSave[iGrp].iDebugVelmpm_AxisA_Uw;    								(*放料A轴调试速度*)
	i_pstStParam_Diamonds_WrRd^.aiDebugGirthmm_AxisA_Uw[iGrp]    		 	:= i_pstStSysParam^.astStGrpParam_UnSave[iGrp].iDebugGirthmm_AxisA_Uw;  								(*放料A轴调试周长*)
//	i_pstStParam_Diamonds_WrRd^.arDebugCurVelmpmAxisA_Uw[iGrp]    		 	:= i_pstStSysParam^.astStGrpParam_UnSave[iGrp].rDebugCurVelmpmAxisA_Uw;  								(*放料A轴调试周长*)
	i_pstStParam_Diamonds_WrRd^.aiDebugVelmpm_AxisB_Uw[iGrp]			 	:= i_pstStSysParam^.astStGrpParam_UnSave[iGrp].iDebugVelmpm_AxisB_Uw;    								(*放料A轴调试速度*)
	i_pstStParam_Diamonds_WrRd^.aiDebugGirthmm_AxisB_Uw[iGrp]    		 	:= i_pstStSysParam^.astStGrpParam_UnSave[iGrp].iDebugGirthmm_AxisB_Uw;  								(*放料A轴调试周长*)
//	i_pstStParam_Diamonds_WrRd^.arDebugCurVelmpmAxisB_Uw[iGrp]    		 	:= i_pstStSysParam^.astStGrpParam_UnSave[iGrp].rDebugCurVelmpmAxisB_Uw;								(*放料A轴调试周长*)
	i_pstStParam_Diamonds_WrRd^.aiDebugVelmpm_AxisA_Rw[iGrp]			 	:= i_pstStSysParam^.astStGrpParam_UnSave[iGrp].iDebugVelmpm_AxisA_Rw;									(*放料A轴调试速度*)
	i_pstStParam_Diamonds_WrRd^.aiDebugGirthmm_AxisA_Rw[iGrp]    		 	:= i_pstStSysParam^.astStGrpParam_UnSave[iGrp].iDebugGirthmm_AxisA_Rw;  								(*放料A轴调试周长*)
//	i_pstStParam_Diamonds_WrRd^.arDebugCurVelmpmAxisA_Rw[iGrp]    		 	:= i_pstStSysParam^.astStGrpParam_UnSave[iGrp].rDebugCurVelmpmAxisA_Rw;								(*放料A轴调试周长*)
	i_pstStParam_Diamonds_WrRd^.aiDebugVelmpm_AxisB_Rw[iGrp]			 	:= i_pstStSysParam^.astStGrpParam_UnSave[iGrp].iDebugVelmpm_AxisB_Rw;									(*放料A轴调试速度*)
	i_pstStParam_Diamonds_WrRd^.aiDebugGirthmm_AxisB_Rw[iGrp]    		 	:= i_pstStSysParam^.astStGrpParam_UnSave[iGrp].iDebugGirthmm_AxisB_Rw;  								(*放料A轴调试周长*)
//	i_pstStParam_Diamonds_WrRd^.arDebugCurVelmpmAxisB_Rw[iGrp]    		 	:= i_pstStSysParam^.astStGrpParam_UnSave[iGrp].rDebugCurVelmpmAxisB_Rw;								(*放料A轴调试周长*)
	i_pstStParam_Diamonds_WrRd^.arVel_Ink[iGrp]							 	:= i_pstStSysParam^.astStGrpParam_Save[iGrp].rVel_Ink;				 								(*空转速度*)
	i_pstStParam_Diamonds_WrRd^.arVel_Inch[iGrp]                      	 	:= i_pstStSysParam^.astStGrpParam_Save[iGrp].rVel_Inch;				 								(*单运行速度*)
	i_pstStParam_Diamonds_WrRd^.abyDelayTime_PressDneInPrint_If[iGrp] 	 	:= i_pstStSysParam^.astStGrpParam_Save[iGrp].byDelayTime_PressDneInPrint_If;		 				(*放牵压辊延时*)
	i_pstStParam_Diamonds_WrRd^.arVel_Max[iGrp]                       	 	:= i_pstStSysParam^.astStGrpParam_Save[iGrp].rVel_Max;		 										(*最大速度*)
	i_pstStParam_Diamonds_WrRd^.abyMeters_UseFollow_1U_V_UwCut[iGrp]	 	:= i_pstStSysParam^.astStGrpParam_Save[iGrp].byMeters_UseFollow_1U_V_UwCut;		 					(*有效距离*)
	i_pstStParam_Diamonds_WrRd^.arGirth_If[iGrp]                    	 	:= i_pstStSysParam^.astStGrpParam_Save[iGrp].rGirth_If;		 										(*放牵辊周长*)
	i_pstStParam_Diamonds_WrRd^.arGirth_Of[iGrp]                    	 	:= i_pstStSysParam^.astStGrpParam_Save[iGrp].rGirth_Of;				 								(*收牵辊周长*)
	i_pstStParam_Diamonds_WrRd^.aiDelayMsec_RollerPress[iGrp]       	 	:= i_pstStSysParam^.astStGrpParam_Save[iGrp].iDelayMsec_RollerPress;								(*合压时间*)
	i_pstStParam_Diamonds_WrRd^.aiTime_S[iGrp]                      	 	:= i_pstStSysParam^.astStGrpParam_Save[iGrp].iTime_S;												(*S加速时间*)
    i_pstStParam_Diamonds_WrRd^.aiTime_S_End[iGrp]                  	 	:= i_pstStSysParam^.astStGrpParam_Save[iGrp].iTime_S_End;											(*S减速时间*)
    i_pstStParam_Diamonds_WrRd^.abyAxisInitPhaseTypeWhenPreRegister[iGrp] 	:= i_pstStSysParam^.astStGrpParam_Save[iGrp].byAxisInitPhaseTypeWhenPreRegister;              		(*预套准初始位置*)
    i_pstStParam_Diamonds_WrRd^.abyVelLimit_PerCent_IfOf[iGrp]            	:= i_pstStSysParam^.astStGrpParam_Save[iGrp].byVelLimit_PerCent_IfOf;         						(*牵引调制限制值*)
    i_pstStParam_Diamonds_WrRd^.arVel_ManuAdjust[iGrp]                    	:= i_pstStSysParam^.astStGrpParam_Save[iGrp].rVel_ManuAdj_Corse;         							(*手动粗调速度*)
    i_pstStParam_Diamonds_WrRd^.arVel_AutoAdjust[iGrp]                    	:= i_pstStSysParam^.astStGrpParam_Save[iGrp].rVel_AutoAdj;         									(*自动调整速度*)
    i_pstStParam_Diamonds_WrRd^.arVel_RapidAdjust[iGrp]                   	:= i_pstStSysParam^.astStGrpParam_Save[iGrp].rVel_RapidAdj;         								(*快速对版速度*)

	i_pstStParam_Diamonds_WrRd^.arAdjVal_PerTime_Fine[iGrp]   		:= i_pstStSysParam^.astStGrpParam_Save[iGrp].rAdjVal_PerTime_Fine;											(*手动细调调整量*)
	i_pstStParam_Diamonds_WrRd^.arAdjVal_PerTime_Coarse[iGrp] 		:= i_pstStSysParam^.astStGrpParam_Save[iGrp].rAdjVal_PerTime_Coarse;										(*手动粗调调整量*)
	i_pstStParam_Diamonds_WrRd^.arVel_HorzAdjust[iGrp]        		:= i_pstStSysParam^.astStGrpParam_Save[iGrp].rVel_HorzdAdj;													(*横向调整速度*)
	i_pstStParam_Diamonds_WrRd^.arVel_HorzPreRegister[iGrp]   		:= i_pstStSysParam^.astStGrpParam_Save[iGrp].rVel_HorzPreRegister;											(*横向预套准速度*)
	i_pstStParam_Diamonds_WrRd^.auiNum_If[iGrp]               		:= i_pstStSysParam^.astStGrpParam_Save[iGrp].uiNum_If;														(*放牵减速比-电机侧*)
	i_pstStParam_Diamonds_WrRd^.auiDen_If[iGrp]               		:= i_pstStSysParam^.astStGrpParam_Save[iGrp].uiDen_If;														(*放牵减速比-传动侧*)
	i_pstStParam_Diamonds_WrRd^.auiNum_Of[iGrp]               		:= i_pstStSysParam^.astStGrpParam_Save[iGrp].uiNum_Of;														(*收牵减速比-电机侧*)
	i_pstStParam_Diamonds_WrRd^.auiDen_Of[iGrp]               		:= i_pstStSysParam^.astStGrpParam_Save[iGrp].uiDen_Of;														(*收牵减速比-传动侧*)
	i_pstStParam_Diamonds_WrRd^.auiNum_Uw[iGrp]               		:= i_pstStSysParam^.astStGrpParam_Save[iGrp].uiNum_Uw;														(*放料减速比-电机侧*)
	i_pstStParam_Diamonds_WrRd^.auiDen_Uw[iGrp]               		:= i_pstStSysParam^.astStGrpParam_Save[iGrp].uiDen_Uw;														(*放料减速比-传动侧*)
	i_pstStParam_Diamonds_WrRd^.auiNum_Rw[iGrp]               		:= i_pstStSysParam^.astStGrpParam_Save[iGrp].uiNum_Rw;														(*收料减速比-电机侧*)
	i_pstStParam_Diamonds_WrRd^.auiDen_Rw[iGrp]               		:= i_pstStSysParam^.astStGrpParam_Save[iGrp].uiDen_Rw;														(*收料减速比-传动侧*)
	i_pstStParam_Diamonds_WrRd^.auiNum_Pu[iGrp]               		:= i_pstStSysParam^.astStGrpParam_Save[iGrp].uiNum_PrnRoller;												(*色组减速比-电机侧*)
	i_pstStParam_Diamonds_WrRd^.auiDen_Pu[iGrp]               		:= i_pstStSysParam^.astStGrpParam_Save[iGrp].uiDen_PrnRoller;												(*色组减速比-传动侧*)
	(*待补充-开始|2025.08.07.202603*)
	(*增加裁切时间集处理2025.9.11.193948*)
	//2026.05.20.214537 修改为直接赋值
	i_pstStParam_Diamonds_WrRd^.astStTimeSet_DnCut_UpCut_Uw_Hmi[iGrp] :=i_pstStSysParam^.astStGrpParam_UnSave[iGrp].stStTimeSet_DnCut_UpCut_Uw_Hmi;
	//2026.05.21.091401 补充收料
	i_pstStParam_Diamonds_WrRd^.astStTimeSet_DnCut_UpCut_Rw_Hmi[iGrp] :=i_pstStSysParam^.astStGrpParam_UnSave[iGrp].stStTimeSet_DnCut_UpCut_Rw_Hmi;

	i_pstStParam_Diamonds_WrRd^.abyAlarmHold_PreCut_Uw[iGrp]:= 	i_pstStSysParam^.astStGrpParam_Save[iGrp].byAlarmHold_PreCut_Uw;
	(*2025.8.26.143548*)
	Action_Input_WrRd_IOTest_MainDOAO();

	(*待补充-结束|2025.08.07.202615*)
	i_pstStParam_Diamonds_WrRd^.arHz_PreHotAir_ManuallySet[iGrp]:= i_pstStSysParam^.astStGrpParam_Save[iGrp].rHz_PreHotAir_ManuallySet;
	i_pstStParam_Diamonds_WrRd^.arSV_PreHeating[iGrp]:= i_pstStSysParam^.astStGrpParam_Save[iGrp].rSV_PreHeating;
	i_pstStParam_Diamonds_WrRd^.arHz_Scraper_ManuallySet[iGrp]:= i_pstStSysParam^.astStGrpParam_Save[iGrp].rHz_Scraper_ManuallySet;
	i_pstStParam_Diamonds_WrRd^.arCoeff_Scraper_Auto[iGrp]:= i_pstStSysParam^.astStGrpParam_Save[iGrp].rCoeff_Scraper_Auto;
	i_pstStParam_Diamonds_WrRd^.arHz_InkRoller_ManuallySet[iGrp]:= i_pstStSysParam^.astStGrpParam_Save[iGrp].rHz_InkRoller_ManuallySet;
	i_pstStParam_Diamonds_WrRd^.arCoeff_InkRoller_Auto[iGrp]:= i_pstStSysParam^.astStGrpParam_Save[iGrp].rCoeff_InkRoller;

	i_pstStParam_Diamonds_WrRd^.auiPreStopDelayTime_ms[iGrp]    := i_pstStSysParam^.astStGrpParam_Save[iGrp].uiPreStopDelayTime_ms	;
	i_pstStParam_Diamonds_WrRd^.arVel_Tar_9905[iGrp]            := i_pstStSysParam^.astStGrpParam_Save[iGrp].rVel_Tar_9905			;
	i_pstStParam_Diamonds_WrRd^.aiAxisId_StepTest_V[iGrp]       := i_pstStSysParam^.astStGrpParam_UnSave[iGrp].iAxisId_StepTest_V		;
	i_pstStParam_Diamonds_WrRd^.aiInterval_StepTest12[iGrp]     := i_pstStSysParam^.astStGrpParam_UnSave[iGrp].iInterval_StepTest12	;
	i_pstStParam_Diamonds_WrRd^.aiMicron_StepTest1_V[iGrp]      := i_pstStSysParam^.astStGrpParam_Save[iGrp].iMicron_StepTest1_V	;
	i_pstStParam_Diamonds_WrRd^.aiMicron_StepTest2_V[iGrp]      := i_pstStSysParam^.astStGrpParam_Save[iGrp].iMicron_StepTest2_V	;
	i_pstStParam_Diamonds_WrRd^.abyKalmanFilterType_Rw[iGrp]    := i_pstStSysParam^.astStGrpParam_Save[iGrp].byKalmanFilterType_Rw	;
	i_pstStParam_Diamonds_WrRd^.abyStructParanInitEn_Rw[iGrp]   := i_pstStSysParam^.astStGrpParam_Save[iGrp].byStructParanInitEn_Rw;

	i_pstStParam_Diamonds_WrRd^.arR_K_MinBeat_Rw[iGrp]          := i_pstStSysParam^.astStGrpParam_Save[iGrp].rR_K_MinBeat_Rw	   ;
	i_pstStParam_Diamonds_WrRd^.aiN_MinBeat_Rw[iGrp]            := i_pstStSysParam^.astStGrpParam_Save[iGrp].iN_MinBeat_Rw	       ;
	i_pstStParam_Diamonds_WrRd^.arR_K_LQR_Rw[iGrp]              := i_pstStSysParam^.astStGrpParam_Save[iGrp].rR_K_LQR_Rw	       ;

	i_pstStParam_Diamonds_WrRd^.arN_LQR_Rw[iGrp]	               	:= i_pstStSysParam^.astStGrpParam_Save[iGrp].rN_LQR_Rw	            ;
	i_pstStParam_Diamonds_WrRd^.arKc_Rw[iGrp]	                   	:= i_pstStSysParam^.astStGrpParam_Save[iGrp].rKc_Rw	            ;
	i_pstStParam_Diamonds_WrRd^.arKc_Rw_AccDec[iGrp]	           	:= i_pstStSysParam^.astStGrpParam_Save[iGrp].rKc_Rw_AccDec	        ;
	i_pstStParam_Diamonds_WrRd^.arWc_LowPass_Diam_Rw[iGrp]	   		:= i_pstStSysParam^.astStGrpParam_Save[iGrp].rWc_LowPass_Diam_Rw	;
	i_pstStParam_Diamonds_WrRd^.abyKalmanFilterType_Uw[iGrp] 	   	:= i_pstStSysParam^.astStGrpParam_Save[iGrp].byKalmanFilterType_Uw ;
	i_pstStParam_Diamonds_WrRd^.abyStructParanInitEn_Uw[iGrp]	   	:= i_pstStSysParam^.astStGrpParam_Save[iGrp].byStructParanInitEn_Uw;

	SysMemCpy(
		ADR(i_pstStParam_Diamonds_WrRd^.astModelParam_Uw[iGrp]),
		ADR(i_pstStSysParam^.astStGrpParam_Save[iGrp].stModelParam_Uw),
		SIZEOF(i_pstStSysParam^.astStGrpParam_Save[iGrp].stModelParam_Uw));
	SysMemCpy(
		ADR(i_pstStParam_Diamonds_WrRd^.astInvariant_Parameters_Uw[iGrp]),
		ADR(i_pstStSysParam^.astStGrpParam_Save[iGrp].stInvariant_Parameters_Uw),
		SIZEOF(i_pstStSysParam^.astStGrpParam_Save[iGrp].stInvariant_Parameters_Uw));
	SysMemCpy(
		ADR(i_pstStParam_Diamonds_WrRd^.astPI_Parameters_Uw[iGrp]),
		ADR(i_pstStSysParam^.astStGrpParam_Save[iGrp].stPI_Parameters_Uw),
		SIZEOF(i_pstStSysParam^.astStGrpParam_Save[iGrp].stPI_Parameters_Uw));
	SysMemCpy(
		ADR(i_pstStParam_Diamonds_WrRd^.astPI_Parameters_Uw_AccDec[iGrp]),
		ADR(i_pstStSysParam^.astStGrpParam_Save[iGrp].stPI_Parameters_Uw_AccDec),
		SIZEOF(i_pstStSysParam^.astStGrpParam_Save[iGrp].stPI_Parameters_Uw_AccDec));

	SysMemCpy(
		ADR(i_pstStParam_Diamonds_WrRd^.astModelParam_Rw[iGrp]),
		ADR(i_pstStSysParam^.astStGrpParam_Save[iGrp].stModelParam_Rw),
		SIZEOF(i_pstStSysParam^.astStGrpParam_Save[iGrp].stModelParam_Rw));
	SysMemCpy(
		ADR(i_pstStParam_Diamonds_WrRd^.astInvariant_Parameters_Rw[iGrp]),
		ADR(i_pstStSysParam^.astStGrpParam_Save[iGrp].stInvariant_Parameters_Rw),
		SIZEOF(i_pstStSysParam^.astStGrpParam_Save[iGrp].stInvariant_Parameters_Rw));
	SysMemCpy(
		ADR(i_pstStParam_Diamonds_WrRd^.astPI_Parameters_Rw[iGrp]),
		ADR(i_pstStSysParam^.astStGrpParam_Save[iGrp].stPI_Parameters_Rw),
		SIZEOF(i_pstStSysParam^.astStGrpParam_Save[iGrp].stPI_Parameters_Rw));
	SysMemCpy(
		ADR(i_pstStParam_Diamonds_WrRd^.astPI_Parameters_Rw_AccDec[iGrp]),
		ADR(i_pstStSysParam^.astStGrpParam_Save[iGrp].stPI_Parameters_Rw_AccDec),
		SIZEOF(i_pstStSysParam^.astStGrpParam_Save[iGrp].stPI_Parameters_Rw_AccDec));

	i_pstStParam_Diamonds_WrRd^.arR_K_MinBeat_Uw[iGrp]    			:= i_pstStSysParam^.astStGrpParam_Save[iGrp].rR_K_MinBeat_Uw    	;
	i_pstStParam_Diamonds_WrRd^.aiN_MinBeat_Uw[iGrp]      			:= i_pstStSysParam^.astStGrpParam_Save[iGrp].iN_MinBeat_Uw      	;
	i_pstStParam_Diamonds_WrRd^.arR_K_LQR_Uw[iGrp]        			:= i_pstStSysParam^.astStGrpParam_Save[iGrp].rR_K_LQR_Uw        	;
	i_pstStParam_Diamonds_WrRd^.arN_LQR_Uw[iGrp]          			:= i_pstStSysParam^.astStGrpParam_Save[iGrp].rN_LQR_Uw          	;
	i_pstStParam_Diamonds_WrRd^.arKc_Uw[iGrp]             			:= i_pstStSysParam^.astStGrpParam_Save[iGrp].rKc_Uw             	;
	i_pstStParam_Diamonds_WrRd^.arKc_Uw_AccDec[iGrp]      			:= i_pstStSysParam^.astStGrpParam_Save[iGrp].rKc_Uw_AccDec      	;
	i_pstStParam_Diamonds_WrRd^.arWc_LowPass_Diam_Uw[iGrp]			:= i_pstStSysParam^.astStGrpParam_Save[iGrp].rWc_LowPass_Diam_Uw	;

	i_pstStParam_Diamonds_WrRd^.arWn_Uw[iGrp]         	      		:= i_pstStSysParam^.astStGrpParam_Save[iGrp].rWn_Uw         	;
	i_pstStParam_Diamonds_WrRd^.arBw_Uw[iGrp]         	      		:= i_pstStSysParam^.astStGrpParam_Save[iGrp].rBw_Uw         	;
	i_pstStParam_Diamonds_WrRd^.arDp_Uw[iGrp]         	      		:= i_pstStSysParam^.astStGrpParam_Save[iGrp].rDp_Uw         	;
	i_pstStParam_Diamonds_WrRd^.aiWorkMode_Pid[iGrp]		  		:= i_pstStSysParam^.astStGrpParam_Save[iGrp].iWorkMode_Pid		;
	i_pstStParam_Diamonds_WrRd^.arFilmLenth_InUnit[iGrp]	   		:= i_pstStSysParam^.astStGrpParam_Save[iGrp].rFilmLenth_InUnit  ;
	i_pstStParam_Diamonds_WrRd^.arTaper_Begin_If[iGrp]:= i_pstStSysParam^.astStGrpParam_Save[iGrp].rTaper_Begin_If;
	i_pstStParam_Diamonds_WrRd^.arTaper_End_If[iGrp]:= i_pstStSysParam^.astStGrpParam_Save[iGrp].rTaper_End_If;
	i_pstStParam_Diamonds_WrRd^.arTaper_Begin_Of[iGrp]:= i_pstStSysParam^.astStGrpParam_Save[iGrp].rTaper_Begin_Of;
	i_pstStParam_Diamonds_WrRd^.arTaper_End_Of[iGrp]:= i_pstStSysParam^.astStGrpParam_Save[iGrp].rTaper_End_Of;
	i_pstStParam_Diamonds_WrRd^.arTaper_Begin_Uw[iGrp]:= i_pstStSysParam^.astStGrpParam_Save[iGrp].rTaper_Begin_Uw;
	i_pstStParam_Diamonds_WrRd^.arTaper_End_Uw[iGrp]:= i_pstStSysParam^.astStGrpParam_Save[iGrp].rTaper_End_Uw;
//2026.1.6.095943增加一些变量
	i_pstStParam_Diamonds_WrRd^.arLength_Band_Confirm[iGrp]:= i_pstStSysParam^.astStGrpParam_Save[iGrp].rLength_Band_Confirm;
	i_pstStParam_Diamonds_WrRd^.arPressure_Tar[iGrp]:= i_pstStSysParam^.astStGrpParam_Save[iGrp].rPressure_Tar;
// 	xSwitch_TensionAdjust_QH					: BIT;
// 	xSwitch_PrnLenAdj_Follow_QH					: BIT;
	i_pstStParam_Diamonds_WrRd^.astBitStWrRd_Switch_Grp[iGrp].xSwitch_TensionAdjust_QH:= i_pstStSysParam^.stStSysParam_Save.dwCtlSwitchRef.3;
	i_pstStParam_Diamonds_WrRd^.astBitStWrRd_Switch_Grp[iGrp].xSwitch_PrnLenAdj_Follow_QH:= i_pstStSysParam^.stStSysParam_Save.dwCtlSwitchRef.2;

	//2026.2.2.165944||新增界面的一些内容|Niu/j
	i_pstStParam_Diamonds_WrRd^.arScrewPitch_PrnRoller_Pressure[iGrp]:= i_pstStSysParam^.astStGrpParam_Save[iGrp].rScrewPitch_PrnRoller_Pressure;
	i_pstStParam_Diamonds_WrRd^.auiNum_PrnRoller_Pressure[iGrp]:= i_pstStSysParam^.astStGrpParam_Save[iGrp].uiNum_PrnRoller_Pressure;
	i_pstStParam_Diamonds_WrRd^.auiDen_PrnRoller_Pressure[iGrp]:= i_pstStSysParam^.astStGrpParam_Save[iGrp].uiDen_PrnRoller_Pressure;

	i_pstStParam_Diamonds_WrRd^.arScrewPitch_NetRoller_Pressure[iGrp]:= i_pstStSysParam^.astStGrpParam_Save[iGrp].rScrewPitch_NetRoller_Pressure;
	i_pstStParam_Diamonds_WrRd^.auiNum_NetRoller_Pressure[iGrp]:= i_pstStSysParam^.astStGrpParam_Save[iGrp].uiNum_NetRoller_Pressure;
	i_pstStParam_Diamonds_WrRd^.auiDen_NetRoller_Pressure[iGrp]:= i_pstStSysParam^.astStGrpParam_Save[iGrp].uiDen_NetRoller_Pressure;

	i_pstStParam_Diamonds_WrRd^.arScrewPitch_StrRoller_Pressure[iGrp]:= i_pstStSysParam^.astStGrpParam_Save[iGrp].rScrewPitch_StrRoller_Pressure;
	i_pstStParam_Diamonds_WrRd^.auiNum_StrRoller_Pressure[iGrp]:= i_pstStSysParam^.astStGrpParam_Save[iGrp].uiNum_StrRoller_Pressure;
	i_pstStParam_Diamonds_WrRd^.auiDen_StrRoller_Pressure[iGrp]:= i_pstStSysParam^.astStGrpParam_Save[iGrp].uiDen_StrRoller_Pressure;

	i_pstStParam_Diamonds_WrRd^.arScrewPitch_Horz[iGrp]:= i_pstStSysParam^.astStGrpParam_Save[iGrp].rScrewPitch_Horz;
	i_pstStParam_Diamonds_WrRd^.auiNum_Horz[iGrp]:= i_pstStSysParam^.astStGrpParam_Save[iGrp].uiNum_Horz;
	i_pstStParam_Diamonds_WrRd^.auiDen_Horz[iGrp]:= i_pstStSysParam^.astStGrpParam_Save[iGrp].uiDen_Horz;

	i_pstStParam_Diamonds_WrRd^.arVel_UVstartVel[iGrp]:= i_pstStSysParam^.astStRSV_GrpParam_Save[iGrp].rVel_UVstartVel;

	//2026.02.28.144731 | + | 上下裁切换
	i_pstStParam_Diamonds_WrRd^.astBitStWrRd_Switch_Grp[iGrp].xSwitch_Change_CutterOnTop_HMI_Uw	:= i_pstStSysParam^.astStGrpParam_Save[iGrp].xSwitch_Change_CutterOnTop_HMI_Uw;(*上下裁切换*)
	i_pstStParam_Diamonds_WrRd^.astBitStWrRd_Switch_Grp[iGrp].xSwitch_Change_CutterOnTop_HMI_Rw	:= i_pstStSysParam^.astStGrpParam_Save[iGrp].xSwitch_Change_CutterOnTop_HMI_Rw;(*上下裁切换*)

	//2026.03.11.100402 | + | 使用Bit22作为压力电机自动合压开关
	i_pstStParam_Diamonds_WrRd^.astBitStWrRd_Switch_Grp[iGrp].xSwitch_PressureAuto_Up_Dn := i_pstStSysParam^.astStGrpParam_Save[iGrp].wCtl_Pressure_Up_Dn.0;

	//2026.03.11.114928 | + | 使用Bit24作为停机维持使能的开关
	i_pstStParam_Diamonds_WrRd^.astBitStWrRd_Switch_Grp[iGrp].xSwitch_KeepServoOn:= i_pstStSysParam^.astStGrpParam_Save[iGrp].dwExtBitCtlFlag.21;

	//2026.02.25.095548 | + | 使用bit23作为天枢数据保存的开关
	i_pstStParam_Diamonds_WrRd^.astBitStWrRd_Switch_Grp[iGrp].xSwitch_SaveData_GNS:= i_pstStSysParam^.astStGrpParam_Save[iGrp].dwExtBitCtlFlag.22;
//2026.04.01.165429 增加总匀墨 Hou.N
	i_pstStParam_Diamonds_WrRd^.astBitStWrRd_Switch_Grp[iGrp].xSwitch_GrpInkEn:=i_pstStSysParam^.astStRSV_GrpParam_UnSave[iGrp].xSwitch_GrpInkEn;

//增加全自动套印相关变量的通讯；2026.4.6.112942|niu.j
	i_pstStParam_Diamonds_WrRd^.astBitStWrRd_Switch_Grp[iGrp].xSwitch_StartAutoFind:= i_pstStSysParam^.astStRSV_GrpParam_UnSave[iGrp].xStartAutoFind;
//增加全自动套印相关变量的通讯；2026.4.6.112942|niu.j
	i_pstStParam_Diamonds_WrRd^.astBitStWrRd_Switch_Grp[iGrp].xSwitch_EnFastPress:= i_pstStSysParam^.astStRSV_GrpParam_Save[iGrp].xSwitch_EnFastPress;
	i_pstStParam_Diamonds_WrRd^.astBitStWrRd_Switch_Grp[iGrp].xSwitch_SaveRS2file:= i_pstStSysParam^.astStRSV_GrpParam_UnSave[iGrp].xSwitch_SaveRS2file;
	i_pstStParam_Diamonds_WrRd^.astBitStWrRd_Switch_Grp[iGrp].xSwitch_RFailure:= i_pstStSysParam^.astStRSV_GrpParam_UnSave[iGrp].xSwitch_RFailure;
	i_pstStParam_Diamonds_WrRd^.astBitStWrRd_Switch_Grp[iGrp].xSwitch_RFailure:= i_pstStSysParam^.astStRSV_GrpParam_UnSave[iGrp].xSwitch_RFailure;
	i_pstStParam_Diamonds_WrRd^.arWidth_Mark_Max[iGrp]:= i_pstStSysParam^.astStRSV_GrpParam_Save[iGrp].rWidth_Mark_Max;
	i_pstStParam_Diamonds_WrRd^.arWidth_Mark_Min[iGrp]:= i_pstStSysParam^.astStRSV_GrpParam_Save[iGrp].rWidth_Mark_Min;
	i_pstStParam_Diamonds_WrRd^.arMaxGap[iGrp]:= i_pstStSysParam^.astStRSV_GrpParam_Save[iGrp].rMaxGap;
	i_pstStParam_Diamonds_WrRd^.arSimilarityThreshold[iGrp]:= i_pstStSysParam^.astStRSV_GrpParam_Save[iGrp].bySimilarityThreshold;
	i_pstStParam_Diamonds_WrRd^.abyMeanOffset[iGrp]:= i_pstStSysParam^.astStRSV_GrpParam_Save[iGrp].byMeanOffset;
	i_pstStParam_Diamonds_WrRd^.abySignalType[iGrp]:= i_pstStSysParam^.astStRSV_GrpParam_Save[iGrp].bySignalType;
	i_pstStParam_Diamonds_WrRd^.arOuterCoff[iGrp]:= i_pstStSysParam^.astStRSV_GrpParam_Save[iGrp].rOuterCoff;
	i_pstStParam_Diamonds_WrRd^.arInnerCoff[iGrp]:= i_pstStSysParam^.astStRSV_GrpParam_Save[iGrp].rInnerCoff;
	FOR iK:=1 TO 15 BY 1 DO
		IF iK<=2 THEN
			i_pstStParam_Diamonds_WrRd^.arFiberMove[iGrp,iK]:= i_pstStSysParam^.astStRSV_GrpParam_Save[iGrp].arFiberMove[iK];
		END_IF
		i_pstStParam_Diamonds_WrRd^.arModeMsg[iGrp,iK]:= i_pstStSysParam^.astStRSV_GrpParam_Save[iGrp].arModeMsg[iK];
	END_FOR

//2026.04.10.234645
	i_pstStParam_Diamonds_WrRd^.abyClrPrnLenCount[iGrp,1]:= i_pstStSysParam^.astStGrpParam_UnSave[iGrp].abyClrPrnLenCount_Rw[1];
	i_pstStParam_Diamonds_WrRd^.abyClrPrnLenCount[iGrp,2]:= i_pstStSysParam^.astStGrpParam_UnSave[iGrp].abyClrPrnLenCount_Rw[2];
	i_pstStParam_Diamonds_WrRd^.abyClrPrnLenCount[iGrp,3]:= i_pstStSysParam^.astStGrpParam_UnSave[iGrp].abyClrPrnLenCount_Rw[3];

//2026.5.12.161016增加速度规划方式的通讯
	i_pstStParam_Diamonds_WrRd^.abyAutoAccDecCurve[iGrp]:= i_pstStSysParam^.astStGrpParam_Save[iGrp].byAutoAccDecCurve;
//2026.05.14.151130 新增自动停机、网辊离压速度
  	i_pstStParam_Diamonds_WrRd^.arRemainDia_stop[iGrp]:=  i_pstStSysParam^.astStRSV_GrpParam_Save[iGrp].rRemainDia_stop  ;
    i_pstStParam_Diamonds_WrRd^.arMaxErr_GantryTrap[iGrp]:= i_pstStSysParam^.astStRSV_GrpParam_Save[iGrp].rMaxErr_GantryTrap ;
    i_pstStParam_Diamonds_WrRd^.arVel_NetReturn[iGrp]:=    i_pstStSysParam^.astStGrpParam_Save[iGrp].rVel_NetReturn ;
    i_pstStParam_Diamonds_WrRd^.astBitStWrRd_Switch_Grp[iGrp].xSwitch_En_AutoStop:=	i_pstStSysParam^.astStRSV_GrpParam_Save[iGrp].xIsAutoStop ;
//2026.05.15.85256 新增电晕启动速度
	i_pstStParam_Diamonds_WrRd^.arVel_CoronaVel[iGrp]:= i_pstStSysParam^.astStRSV_GrpParam_Save[iGrp].rVel_CoronaVel;
	(*2026.05.26.155311+*)
	i_pstStParam_Diamonds_WrRd^.astBitStWrRd_Switch_Grp[iGrp].xAutoAccDec_Hmi:=	i_pstStSysParam^.astStGrpParam_UnSave[iGrp].xAutoAccDec_Hmi ;

//2026.05.24.135821 光纤行走部分
	i_pstStParam_Diamonds_WrRd^.aiFiberMoveVel[iGrp]:= i_pstStSysParam^.astStRSV_GrpParam_Save[iGrp].iFiberMoveVel;
	i_pstStParam_Diamonds_WrRd^.arFiberMoveDistance_AllUnit[iGrp]:= i_pstStSysParam^.astStRSV_GrpParam_UnSave[iGrp].rFiberMoveDistance_AllUnit;
	i_pstStParam_Diamonds_WrRd^.abyFiberMove_MicroMoveStep[iGrp]:= i_pstStSysParam^.astStRSV_GrpParam_Save[iGrp].byFiberMove_MicroMoveStep;
	i_pstStParam_Diamonds_WrRd^.astBitStWrRd_Switch_Grp[iGrp].xFiberMove_DebugMode:=i_pstStSysParam^.astStRSV_GrpParam_UnSave[iGrp].xFiberMove_DebugMode;
	i_pstStParam_Diamonds_WrRd^.astBitStWrRd_Switch_Grp[iGrp].xFiberMoveDisRunStart_AllUnit:=i_pstStSysParam^.astStRSV_GrpParam_UnSave[iGrp].xFiberMoveDisRunStart_AllUnit;
	i_pstStParam_Diamonds_WrRd^.astBitStWrRd_Switch_Grp[iGrp].xUseOnline_FiberMove:=i_pstStSysParam^.astStRSV_GrpParam_Save[iGrp].xUseOnline_FiberMove;
	i_pstStParam_Diamonds_WrRd^.astBitStWrRd_Switch_Grp[iGrp].xFiberMoveConfirm_AllUnit:=i_pstStSysParam^.astStRSV_GrpParam_UnSave[iGrp].xFiberMoveConfirm_AllUnit;
	i_pstStParam_Diamonds_WrRd^.astBitStWrRd_Switch_Grp[iGrp].xFiberMovePosCal_ByUnit:=i_pstStSysParam^.astStRSV_GrpParam_UnSave[iGrp].xFiberMovePosCal_ByUnit;
	i_pstStParam_Diamonds_WrRd^.astBitStWrRd_Switch_Grp[iGrp].xFiberMovePosCal_ByOnline:=i_pstStSysParam^.astStRSV_GrpParam_UnSave[iGrp].xFiberMovePosCal_ByOnline;
	i_pstStParam_Diamonds_WrRd^.astBitStWrRd_Switch_Grp[iGrp].xFiberMove_Negative_AdjustByUnit:=i_pstStSysParam^.astStRSV_GrpParam_Save[iGrp].xFiberMove_Negative_AdjustByUnit;
	i_pstStParam_Diamonds_WrRd^.astBitStWrRd_Switch_Grp[iGrp].xFiberMove_Negative_AdjustByOnline:=i_pstStSysParam^.astStRSV_GrpParam_Save[iGrp].xFiberMove_Negative_AdjustByOnline;
//2026.5.15.112026增加卷径检测变量输入
	FOR iK:=1 TO 4 BY 1 DO
		i_pstStParam_Diamonds_WrRd^.arStdVol_Coef_Axis_Hmi[iGrp,iK]:= i_pstStSysParam^.astStGrpParam_UnSave[iGrp].alrStdVol_Coef_Axis_Hmi[iK];
		i_pstStParam_Diamonds_WrRd^.arStdVol_Diam_Axis_Hmi[iGrp,iK]:= i_pstStSysParam^.astStGrpParam_UnSave[iGrp].alrStdVol_Diam_Axis_Hmi[iK];
		i_pstStParam_Diamonds_WrRd^.arStdVol_Volt_Axis_Hmi[iGrp,iK]:= i_pstStSysParam^.astStGrpParam_UnSave[iGrp].alrStdVol_Volt_Axis_Hmi[iK];
	END_FOR
	i_pstStParam_Diamonds_WrRd^.arStdVol_Coef_Axis_Hmi[iGrp,0]:= i_pstStSysParam^.astStGrpParam_UnSave[iGrp].alrStdVol_Coef_Axis_Hmi[0];

END_FOR
(*轴参数|2025.08.07.101610*)
FOR iUnitId:= 1 TO MAX_UNIT_NUM BY 1 DO
	(*待补充-开始|2025.08.07.112308*)

	i_pstStParam_Diamonds_WrRd^.astStWrRd_UnitParam[iUnitId].stBitStWrRd_Switch_Unit.xSwitch_CoatingPrn					:= i_pstStSysParam^.astStUnitParam_Save[iUnitId].xSwitchOn_CoatingPrn ;(*色组涂布开关*)
	i_pstStParam_Diamonds_WrRd^.astStWrRd_UnitParam[iUnitId].stBitStWrRd_Switch_Unit.xSwitch_CoatingRec					:= i_pstStSysParam^.astStUnitParam_Save[iUnitId].xReverseAdj_CoatingPrn ;(*涂布调整反向*)
	i_pstStParam_Diamonds_WrRd^.astStWrRd_UnitParam[iUnitId].stBitStWrRd_Switch_Unit.xSwitch_ScraperAuto				:= i_pstStSysParam^.astStUnitParam_Save[iUnitId].xSwitch_ScraperAuto ;(*刮刀手自动*)
	i_pstStParam_Diamonds_WrRd^.astStWrRd_UnitParam[iUnitId].stBitStWrRd_Switch_Unit.xSwitch_ScraperOn					:= i_pstStSysParam^.astStUnitParam_Save[iUnitId].xSwitch_ScraperOn ;(*刮刀开关*)
	i_pstStParam_Diamonds_WrRd^.astStWrRd_UnitParam[iUnitId].stBitStWrRd_Switch_Unit.xSwitch_InkRollerAuto				:= i_pstStSysParam^.astStUnitParam_Save[iUnitId].xSwitch_InkRollerAuto ;(*递墨辊手自动*)
	i_pstStParam_Diamonds_WrRd^.astStWrRd_UnitParam[iUnitId].stBitStWrRd_Switch_Unit.xSwitch_InkRollerCW				:= i_pstStSysParam^.astStUnitParam_Save[iUnitId].xSwitch_InkRollerCW ;(*递墨辊正转*)
	i_pstStParam_Diamonds_WrRd^.astStWrRd_UnitParam[iUnitId].stBitStWrRd_Switch_Unit.xSwitch_InkRollerCCW				:= i_pstStSysParam^.astStUnitParam_Save[iUnitId].xSwitch_InkRollerCCW ;(*递墨辊反转*)
	i_pstStParam_Diamonds_WrRd^.astStWrRd_UnitParam[iUnitId].stBitStWrRd_Switch_Unit.xSwitch_HotWindOn					:= i_pstStSysParam^.astStUnitParam_Save[iUnitId].xSwitch_HotWindOn ;(*热风开关*)
//	i_pstStParam_Diamonds_WrRd^.astStWrRd_UnitParam[iUnitId].stBitStWrRd_Switch_Unit.xSwitch_HeatingOn					:= i_pstStSysParam^.astStUnitParam_Save[iUnitId].xSwitch_HeatingOn ;(*加热开关*)
	i_pstStParam_Diamonds_WrRd^.astStWrRd_UnitParam[iUnitId].stBitStWrRd_Switch_Unit.xSwitch_Heating_I					:= i_pstStSysParam^.astStUnitParam_Save[iUnitId].xSwitch_Heating_I ;(*加热I档*)
	i_pstStParam_Diamonds_WrRd^.astStWrRd_UnitParam[iUnitId].stBitStWrRd_Switch_Unit.xSwitch_Heating_II					:= i_pstStSysParam^.astStUnitParam_Save[iUnitId].xSwitch_Heating_II ;(*加热II档*)
	i_pstStParam_Diamonds_WrRd^.astStWrRd_UnitParam[iUnitId].stBitStWrRd_Switch_Unit.xSwitch_Heating_III				:= i_pstStSysParam^.astStUnitParam_Save[iUnitId].xSwitch_Heating_III ;(*加热III档*)
	i_pstStParam_Diamonds_WrRd^.astStWrRd_UnitParam[iUnitId].stBitStWrRd_Switch_Unit.xSwitch_ThisUnitEna				:= i_pstStSysParam^.astStUnitParam_Save[iUnitId].xEnable_arc ;(*色组套印开关*)
	i_pstStParam_Diamonds_WrRd^.astStWrRd_UnitParam[iUnitId].stBitStWrRd_Switch_Unit.xSwitch_Horz						:= i_pstStSysParam^.astStUnitParam_Save[iUnitId].dwFlag_Ctl.0 ;(*横向开关*)
	i_pstStParam_Diamonds_WrRd^.astStWrRd_UnitParam[iUnitId].stBitStWrRd_Switch_Unit.xSwitch_DoorBaseLn					:= i_pstStSysParam^.astStUnitParam_Save[iUnitId].dwFlag_Ctl.1 ;(*门内基线开关*)
//	i_pstStParam_Diamonds_WrRd^.astStWrRd_UnitParam[iUnitId].stBitStWrRd_Switch_Unit.xSwitch_SmallSignalProcessing_T1_1	:= i_pstStSysParam^.astStUnitParam_Save[iUnitId]. ;(*第一组波门T1内小信号处理开关*)
//	i_pstStParam_Diamonds_WrRd^.astStWrRd_UnitParam[iUnitId].stBitStWrRd_Switch_Unit.xSwitch_SmallSignalProcessing_T2_1	:= i_pstStSysParam^.astStUnitParam_Save[iUnitId]. ;(*第一组波门T2内小信号处理开关*)
//	i_pstStParam_Diamonds_WrRd^.astStWrRd_UnitParam[iUnitId].stBitStWrRd_Switch_Unit.xSwitch_SmallSignalProcessing_T1_2	:= i_pstStSysParam^.astStUnitParam_Save[iUnitId]. ;(*第二组波门T1内小信号处理开关*)
//	i_pstStParam_Diamonds_WrRd^.astStWrRd_UnitParam[iUnitId].stBitStWrRd_Switch_Unit.xSwitch_SmallSignalProcessing_T2_2	:= i_pstStSysParam^.astStUnitParam_Save[iUnitId]. ;(*第二组波门T2内小信号处理开关*)
(*小信号2025.10.27.141809*)
	i_pstStParam_Diamonds_WrRd^.astStWrRd_UnitParam[iUnitId].stBitStWrRd_Switch_Unit.xSwitch_SmallSignalProcessing_T1:= i_pstStSysParam^.astStUnitParam_Save[iUnitId].dwFlag_Ctl.13;
	i_pstStParam_Diamonds_WrRd^.astStWrRd_UnitParam[iUnitId].stBitStWrRd_Switch_Unit.xSwitch_SmallSignalProcessing_T2:= i_pstStSysParam^.astStUnitParam_Save[iUnitId].dwFlag_Ctl.14;
